(* CODESYS project Syn_Visu_9.4.0.library
   Version: 9.4.0.0
   Title: SynVisu
   Placeholder: SynVisu
   Company: Syntegon Group
   DefaultNamespace: SynVisu

Project tree, tasks and I/O mapping:
  libraries: Tc2_System, * (Beckhoff Automation GmbH)
  DUTs/
    data type E_VisuBodyRole
    data type E_VisuBodyShape
    data type E_VisuCartesianAxes
    data type E_VisuComponentType
    data type E_VisuModuleKind
    data type E_VisuProductShape
    data type E_VisuProductState
    data type ST_VisuBody
    data type ST_VisuBodyState
    data type ST_VisuCartesian
    data type ST_VisuCartesianConfig
    data type ST_VisuCartesianState
    data type ST_VisuConveyor
    data type ST_VisuConveyorConfig
    data type ST_VisuConveyorState
    data type ST_VisuDelta
    data type ST_VisuDeltaConfig
    data type ST_VisuDeltaState
    data type ST_VisuDetector
    data type ST_VisuDetectorConfig
    data type ST_VisuDetectorState
    data type ST_VisuFault
    data type ST_VisuFinger
    data type ST_VisuFingerState
    data type ST_VisuGantryMover
    data type ST_VisuLimitArea
    data type ST_VisuLoopMover
    data type ST_VisuManifest
    data type ST_VisuManifestEntry
    data type ST_VisuPlanarPose
    data type ST_VisuPose
    data type ST_VisuPosition
    data type ST_VisuProduct
    data type ST_VisuProductType
    data type ST_VisuStation
    data type ST_VisuStationConfig
    data type ST_VisuStationState
    data type ST_VisuTrackModule
    data type ST_VisuTrackModuleState
    data type ST_VisuWorkingArea
    data type ST_VisuXtsGantry
    data type ST_VisuXtsGantryConfig
    data type ST_VisuXtsGantryState
    data type ST_VisuXtsLoop
    data type ST_VisuXtsLoopConfig
    data type ST_VisuXtsLoopState
    data type ST_VisuZone
  GVLs/
    global variables VISU_GlobalConst
    global variables VISU_GlobalConst_Param
  POUs/
    function block _FB_VisuBodyComponent [ST]: m_ClearBodies, m_Parts, m_Register, m_SetBody, m_SetBodyActive, m_SetFault, m_SetOriginShift, m_SetPose
    function block _FB_VisuCartesian [ST]: m_ApplyConfig, m_ComponentType, m_Configure, m_Fingers, m_LimitArea, m_SetAxes, m_SetFault, m_SetFingerState, m_SetKinematics, m_SetOriginShift, m_Zones
    function block _FB_VisuComponent [ST]: m_ComponentType, m_DcTime, m_Id, m_NotifyConfigChanged, m_Register, m_SymbolPath
    function block _FB_VisuConveyor [ST]: m_ApplyConfig, m_BeltPosition, m_ComponentType, m_Configure, m_FindProduct, m_GetProduct, m_IndexInsert, m_IndexRebuild, m_IndexSlotOf, m_LatchProduct, m_MoveProduct, m_ProductCount, m_ProductPose, m_RemoveProduct, m_RemoveProductsBeyond, m_SetBeltPosition, m_SetBodyVisible, m_SetFault, m_SetModuloBeltPosition, m_SetOriginShift, m_SetProductState, m_SetProductType, m_StaysInRegister
    function block _FB_VisuDelta [ST]: m_ApplyConfig, m_BasePose, m_ComponentType, m_Configure, m_Fingers, m_LimitArea, m_SetFault, m_SetFingerState, m_SetOriginShift, m_SetTcp, m_SetWorkingArea, m_Zones
    function block _FB_VisuDetector [ST]: m_Parts, m_Zones
    function block _FB_VisuRobot [ST]: m_ClearFingers, m_ClearLimitArea, m_ClearTcpLimitArea, m_Fingers, m_LimitArea, m_SetFinger, m_SetLimitArea, m_SetTcpLimitArea
    function block _FB_VisuSensor [ST]: m_ComponentType, m_Configure, m_SetSignal
    function block _FB_VisuStation [ST]: m_ComponentType, m_Configure, m_Parts, m_Zones
    function block _FB_VisuVision [ST]: m_ComponentType, m_Configure
    function block _FB_VisuXtsGantry [ST]: m_ApplyConfig, m_ComponentType, m_Configure, m_Fingers, m_LimitArea, m_Modules, m_SetFault, m_SetMover, m_SetMoverCount, m_SetOriginShift, m_SetZPosition, m_Zones
    function block _FB_VisuXtsLoop [ST]: m_ApplyConfig, m_ComponentType, m_Configure, m_Fingers, m_LimitArea, m_Modules, m_SetFault, m_SetMover, m_SetMoverCount, m_SetOriginShift, m_Zones
    function block _FB_VisuXtsTrack [ST]: m_ClearModules, m_Modules, m_SetModule, m_SetModuleFault, m_TrackLength
    function block _FB_VisuZoneComponent [ST]: m_ClearZones, m_SetZone, m_Zones
    function _FC_GetVersionSynVisu [ST]
*)

// DUTs/E_VisuBodyRole
{attribute 'qualified_only'}
{attribute 'strict'}
TYPE E_VisuBodyRole :
(
	(* Values are part of the gateway contract: append, never renumber. What a body stands for sets its look. *)
	STRUCTURE := 0,		// machine part: lit, with shadow
	SENSOR := 1,		// sensing part, e.g. a lens or a light barrier head: lit, in its own colour
	BEAM := 2,			// overlay on the zones layer, lights up while active
	FIELD_OF_VIEW := 3	// overlay on the zones layer, lights up while active
) UINT;
END_TYPE

// DUTs/E_VisuBodyShape
{attribute 'qualified_only'}
{attribute 'strict'}
TYPE E_VisuBodyShape :
(
	(* Values are part of the gateway contract: append, never renumber. *)
	BOX := 0,			// box: fLength x fWidth x fHeight
	CYLINDER := 1,		// cylinder: fLength and fWidth are its two diameters
	FRUSTUM := 2		// rectangular pyramid stump: bottom fLength x fWidth, top fTopLength x fTopWidth
) UINT;
END_TYPE

// DUTs/E_VisuCartesianAxes
{attribute 'qualified_only'}
{attribute 'strict'}
TYPE E_VisuCartesianAxes :
(
	(* Values are part of the gateway contract: append, never renumber. Which axes a Cartesian robot has. *)
	XYZ := 0,	// rails along local Y, bridge (Y), carriage (X) and column (Z)
	XZ := 1,	// no Y axis: a fixed beam along local X at fRailHeight, carriage (X) and column (Z); Y is always 0
	XY := 2		// no Z axis: rails, bridge (Y) and carriage (X); the column has a fixed length, the flange stays at fZMin
) UINT;
END_TYPE

// DUTs/E_VisuComponentType
{attribute 'qualified_only'}
{attribute 'strict'}
TYPE E_VisuComponentType :
(
	(* Values are part of the gateway contract: append, never renumber. *)
	NONE := 0,
	CONVEYOR := 1,
	DELTA := 2,
	XTS_GANTRY := 3,
	XTS_LOOP := 4,
	CARTESIAN := 5,
	VISION := 6,
	SENSOR := 7,
	STATION := 8
) UINT;
END_TYPE

// DUTs/E_VisuModuleKind
{attribute 'qualified_only'}
{attribute 'strict'}
TYPE E_VisuModuleKind :
(
	(* Values are part of the gateway contract: append, never renumber. What an XTS track module is. *)
	STRAIGHT := 0,		// straight motor module
	CURVE_LEFT := 1,	// curve module: turns the track by a quarter circle (90 deg) to the left
	CURVE_RIGHT := 2	// curve module: turns the track by a quarter circle (90 deg) to the right
) UINT;
END_TYPE

// DUTs/E_VisuProductShape
{attribute 'qualified_only'}
{attribute 'strict'}
TYPE E_VisuProductShape :
(
	(* Values are part of the gateway contract: append, never renumber. *)
	BOX := 0,			// box: fLength x fWidth x fHeight
	CYLINDER := 1,		// cylinder: fLength and fWidth are its diameters along and across the conveying direction
	ROUNDED_BOX := 2	// box with rounded vertical edges of fCornerRadius (pouches, flow packs)
) UINT;
END_TYPE

// DUTs/E_VisuProductState
{attribute 'qualified_only'}
{attribute 'strict'}
TYPE E_VisuProductState :
(
	(* Values are part of the gateway contract: append, never renumber. *)
	DETECTED := 0,
	ASSIGNED := 1,
	PICKED := 2,
	REJECTED := 3,
	PLACED := 4
) UINT;
END_TYPE

// DUTs/ST_VisuBody
TYPE ST_VisuBody :
STRUCT
	(* One solid a component is drawn from, so the visualisation needs no code of its own for it. It stands on
	   its bottom face and extends along its local +Z. *)
	eShape : E_VisuBodyShape;
	eRole : E_VisuBodyRole;
	stPose : ST_VisuPose; // bottom centre in the component's frame (from its stPose), not MCS
	fLength : LREAL; // mm along the body's local X
	fWidth : LREAL; // mm along the body's local Y
	fHeight : LREAL; // mm along the body's local Z
	fTopLength : LREAL; // mm, top face of a FRUSTUM
	fTopWidth : LREAL; // mm, top face of a FRUSTUM
END_STRUCT
END_TYPE

// DUTs/ST_VisuBodyState
TYPE ST_VisuBodyState :
STRUCT
	bActive : BOOL; // a BEAM or FIELD_OF_VIEW lights up, e.g. an interrupted light barrier
END_STRUCT
END_TYPE

// DUTs/ST_VisuCartesian
TYPE ST_VisuCartesian :
STRUCT
	(* One visualised Cartesian robot. Register the instance's symbol path in the manifest with
	   eType := E_VisuComponentType.CARTESIAN. *)
	stConfig : ST_VisuCartesianConfig; // read at discovery and after nConfigVersion changes
	stState : ST_VisuCartesianState; // read every gateway cycle
END_STRUCT
END_TYPE

// DUTs/ST_VisuCartesianConfig
TYPE ST_VisuCartesianConfig :
STRUCT
	(* Cartesian robot: two fixed rails along local +Y, a bridge travelling in Y, a carriage on it travelling in X
	   and a vertical column (Z) ending at the gripper flange. Local frame: origin at axis X = Y = 0, Z up; the
	   flange is at (X, Y, Z). Without a Y axis (eAxes XZ) a fixed beam along X at fRailHeight replaces rails and
	   bridge and Y is 0; without a Z axis (XY) the column has a fixed length and the flange stays at fZMin. *)
	stPose : ST_VisuPose; // MCS
	eAxes : E_VisuCartesianAxes := E_VisuCartesianAxes.XYZ; // which axes the robot has (set by m_SetKinematics)
	fXMin : LREAL; // mm, X stroke
	fXMax : LREAL; // mm
	fYMin : LREAL; // mm, Y stroke
	fYMax : LREAL; // mm
	fZMin : LREAL; // mm, Z stroke
	fZMax : LREAL; // mm
	fRailHeight : LREAL; // mm, top of the rails above the local origin; the bridge sits on them
	stLimitArea : ST_VisuLimitArea; // optional box in the robot frame that further restricts the working area
	stTcpLimitArea : ST_VisuLimitArea; // optional box around the gripper flange, along the robot frame's axes
	nZoneCount : UINT;
	aZones : ARRAY[0..VISU_GlobalConst_Param.VISU_un_MAX_ZONES - 1] OF ST_VisuZone; // pick and place zones
	nFingerCount : UINT; // 0 = no gripper definition
	aFingers : ARRAY[0..VISU_GlobalConst_Param.VISU_un_MAX_FINGERS - 1] OF ST_VisuFinger;
	(* mm in the local frame from stPose: origin of the robot's coordinate system as shown (origin triad, local
	   measuring coordinates). The geometry and axis values stay relative to stPose. *)
	stOriginShift : ST_VisuPosition;
END_STRUCT
END_TYPE

// DUTs/ST_VisuCartesianState
TYPE ST_VisuCartesianState :
STRUCT
	nTimestamp : ULINT; // DC time of the writing cycle, ns since 2000-01-01 (set by _FB_VisuCartesian)
	fX : LREAL; // mm, actual value: the gripper flange
	fY : LREAL; // mm, actual value
	fZ : LREAL; // mm, actual value
	bGripperActive : BOOL; // used only when no fingers are configured
	aFingerStates : ARRAY[0..VISU_GlobalConst_Param.VISU_un_MAX_FINGERS - 1] OF ST_VisuFingerState; // one per configured finger
	stFault : ST_VisuFault; // fault of the robot (set by _FB_VisuCartesian.m_SetFault)
END_STRUCT
END_TYPE

// DUTs/ST_VisuConveyor
TYPE ST_VisuConveyor :
STRUCT
	(* One visualised conveyor. Register the instance's symbol path in the manifest with
	   eType := E_VisuComponentType.CONVEYOR. *)
	stConfig : ST_VisuConveyorConfig; // read at discovery and after nConfigVersion changes
	stState : ST_VisuConveyorState; // read every gateway cycle
END_STRUCT
END_TYPE

// DUTs/ST_VisuConveyorConfig
TYPE ST_VisuConveyorConfig :
STRUCT
	stPose : ST_VisuPose; // belt start on the belt surface; local +X = conveying direction
	fLength : LREAL; // mm
	fWidth : LREAL; // mm
	nProductTypeCount : UINT;
	aProductTypes : ARRAY[0..VISU_GlobalConst_Param.VISU_un_MAX_PRODUCT_TYPES - 1] OF ST_VisuProductType;
	bBody : BOOL := TRUE; // TRUE = the belt is drawn as a body; FALSE = a conveyor without one (products, zones and axis only)
	(* mm in the local frame from stPose: origin of the conveyor's coordinate system. Belt coordinates (zones'
	   fStart, fEnd, fCcsOffset) count from this origin. 0 = the belt start. *)
	stOriginShift : ST_VisuPosition;
END_STRUCT
END_TYPE

// DUTs/ST_VisuConveyorState
TYPE ST_VisuConveyorState :
STRUCT
	nTimestamp : ULINT; // DC time of the writing cycle, ns since 2000-01-01 (set by _FB_VisuConveyor)
	fBeltPosition : LREAL; // continuous belt surface position, mm, no modulo (see _FB_VisuConveyor.m_SetModuloBeltPosition)
	nProductCount : UINT; // entries [0..nProductCount-1] are evaluated
	aProducts : ARRAY[0..VISU_GlobalConst_Param.VISU_un_MAX_PRODUCTS - 1] OF ST_VisuProduct;
	stFault : ST_VisuFault; // fault of the conveyor (set by _FB_VisuConveyor.m_SetFault)
END_STRUCT
END_TYPE

// DUTs/ST_VisuDelta
TYPE ST_VisuDelta :
STRUCT
	(* One visualised Delta robot. Register the instance's symbol path in the manifest with
	   eType := E_VisuComponentType.DELTA. *)
	stConfig : ST_VisuDeltaConfig; // read at discovery and after nConfigVersion changes
	stState : ST_VisuDeltaState; // read every gateway cycle
END_STRUCT
END_TYPE

// DUTs/ST_VisuDeltaConfig
TYPE ST_VisuDeltaConfig :
STRUCT
	(* Geometry the visualisation uses to derive the arm posture from the TCP.
	   Arm 1 lies along the base's local +X; arms 2 and 3 follow counter-clockwise
	   (seen from above) at 120 deg each. *)
	stPose : ST_VisuPose; // base centre in the MCS
	fBaseRadius : LREAL; // mm, base centre to shoulder joint
	fEffectorRadius : LREAL; // mm, effector centre to lower-arm joint
	fUpperArmLength : LREAL; // mm
	fLowerArmLength : LREAL; // mm
	stWorkingArea : ST_VisuWorkingArea;
	stLimitArea : ST_VisuLimitArea; // optional box that further restricts the working area
	stTcpLimitArea : ST_VisuLimitArea; // optional box around the TCP, relative to it along the robot frame's axes
	nZoneCount : UINT;
	aZones : ARRAY[0..VISU_GlobalConst_Param.VISU_un_MAX_ZONES - 1] OF ST_VisuZone; // pick and place zones
	nFingerCount : UINT; // 0 = no gripper definition
	aFingers : ARRAY[0..VISU_GlobalConst_Param.VISU_un_MAX_FINGERS - 1] OF ST_VisuFinger;
	(* mm in the local frame from stPose: origin of the robot's coordinate system as shown (origin triad, local
	   measuring coordinates). The geometry, working area and limit area stay relative to stPose. *)
	stOriginShift : ST_VisuPosition;
END_STRUCT
END_TYPE

// DUTs/ST_VisuDeltaState
TYPE ST_VisuDeltaState :
STRUCT
	nTimestamp : ULINT; // DC time of the writing cycle, ns since 2000-01-01 (set by _FB_VisuDelta.m_SetTcp)
	stActualTcp : ST_VisuPosition; // MCS, effector centre (the gripper flange); the visualisation derives the arms from it
	stSetpointTcp : ST_VisuPosition; // MCS
	aFingerStates : ARRAY[0..VISU_GlobalConst_Param.VISU_un_MAX_FINGERS - 1] OF ST_VisuFingerState; // one per configured finger
	stFault : ST_VisuFault; // fault of the robot (set by _FB_VisuDelta.m_SetFault)
END_STRUCT
END_TYPE

// DUTs/ST_VisuDetector
TYPE ST_VisuDetector :
STRUCT
	(* One visualised vision system or product sensor. Register the instance's symbol path in the manifest with
	   eType := E_VisuComponentType.VISION or SENSOR; both share this structure. *)
	stConfig : ST_VisuDetectorConfig; // read at discovery and after nConfigVersion changes
	stState : ST_VisuDetectorState; // read every gateway cycle
END_STRUCT
END_TYPE

// DUTs/ST_VisuDetectorConfig
TYPE ST_VisuDetectorConfig :
STRUCT
	(* A detector (vision system, product sensor): its zones on the conveyors and the bodies it is drawn from. *)
	stPose : ST_VisuPose; // MCS; a vision system's lens looking along local -Z, a sensor's head
	nZoneCount : UINT;
	aZones : ARRAY[0..VISU_GlobalConst_Param.VISU_un_MAX_ZONES - 1] OF ST_VisuZone; // where it detects
	nBodyCount : UINT;
	aBodies : ARRAY[0..VISU_GlobalConst_Param.VISU_un_MAX_BODIES - 1] OF ST_VisuBody;
	(* mm in the local frame from stPose: origin of the detector's coordinate system as shown (origin triad, local
	   measuring coordinates). The bodies stay relative to stPose. *)
	stOriginShift : ST_VisuPosition;
END_STRUCT
END_TYPE

// DUTs/ST_VisuDetectorState
TYPE ST_VisuDetectorState :
STRUCT
	nTimestamp : ULINT; // DC time of the writing cycle, ns since 2000-01-01 (set by _FB_VisuDetector)
	aBodyStates : ARRAY[0..VISU_GlobalConst_Param.VISU_un_MAX_BODIES - 1] OF ST_VisuBodyState; // one per configured body
	stFault : ST_VisuFault; // fault of the detector (set by _FB_VisuDetector.m_SetFault)
END_STRUCT
END_TYPE

// DUTs/ST_VisuFault
(* Fault of a component or an XTS mover: drawn red with sMessage while bActive (contract, protocol 8). *)
TYPE ST_VisuFault :
STRUCT
	bActive : BOOL; // TRUE while the fault is active
	sMessage : STRING(80); // shown to the operator; empty shows 'Fault'
END_STRUCT
END_TYPE

// DUTs/ST_VisuFinger
TYPE ST_VisuFinger :
STRUCT
	(* One gripper finger, always drawn as a cylinder. Its frame's origin is the centre of its top face; it extends
	   along its local -Z. The grip point, where a carried product's top touches, is the centre of its bottom face. *)
	fDiameter : LREAL; // mm
	fHeight : LREAL; // mm
END_STRUCT
END_TYPE

// DUTs/ST_VisuFingerState
TYPE ST_VisuFingerState :
STRUCT
	stPose : ST_VisuPose; // MCS, absolute: pose of the finger's frame (centre of its top face)
	bActive : BOOL; // the finger grips
END_STRUCT
END_TYPE

// DUTs/ST_VisuGantryMover
TYPE ST_VisuGantryMover :
STRUCT
	nId : UDINT; // unique within the gantry, > 0; referenced by a carried product's nMoverId
	bValid : BOOL; // invalid entries are not shown
	fPosition : LREAL; // mm along the track (local +Y), actual value
	fX : LREAL; // mm, X axis on the mover, actual value
	bGripperActive : BOOL; // used only when no fingers are configured
	aFingerStates : ARRAY[0..VISU_GlobalConst_Param.VISU_un_MAX_FINGERS - 1] OF ST_VisuFingerState; // one per configured finger
	stFault : ST_VisuFault; // fault of this mover
END_STRUCT
END_TYPE

// DUTs/ST_VisuLimitArea
TYPE ST_VisuLimitArea :
STRUCT
	(* Axis-aligned box along the robot frame's axes (turned with its stPose). As stLimitArea it lies in the robot
	   frame (relative to stPose, the frame its working area is given in) and further restricts the working area, e.g.
	   so that neighbouring robots cannot collide (_FB_VisuRobot.m_SetLimitArea). As stTcpLimitArea it lies around the
	   TCP (XTS gantry: every mover's gripper flange), relative to it, and moves with it without turning
	   (_FB_VisuRobot.m_SetTcpLimitArea): the visualisation flags it when it overlaps another robot's limit area or
	   TCP limit area or leaves its own robot's limit area. Delta, XTS gantry and Cartesian robot; an XTS loop has
	   neither. *)
	fXMin : LREAL; // mm
	fXMax : LREAL; // mm
	fYMin : LREAL; // mm
	fYMax : LREAL; // mm
	fZMin : LREAL; // mm relative to the base or the TCP (below it: negative)
	fZMax : LREAL; // mm relative to the base or the TCP
	bActive : BOOL; // FALSE: no box, nothing is drawn or checked
END_STRUCT
END_TYPE

// DUTs/ST_VisuLoopMover
TYPE ST_VisuLoopMover :
STRUCT
	nId : UDINT; // unique within the loop, > 0; referenced by a carried product's nMoverId
	bValid : BOOL; // invalid entries are not shown
	fPosition : LREAL; // mm along the loop from the start of the lower straight, in the conveying direction
	aFingerStates : ARRAY[0..VISU_GlobalConst_Param.VISU_un_MAX_FINGERS - 1] OF ST_VisuFingerState; // one per configured finger
	stFault : ST_VisuFault; // fault of this mover
END_STRUCT
END_TYPE

// DUTs/ST_VisuManifest
TYPE ST_VisuManifest :
STRUCT
	(* Discovery entry point. The application declares one instance at the fixed symbol
	   GVL_Visu.stManifest; the gateway starts reading there. *)
	nProtocolVersion : UINT := VISU_GlobalConst.VISU_un_PROTOCOL_VERSION;
	(* Increment after any change to the manifest or to a component's stConfig. *)
	nConfigVersion : UDINT := 1;
	nCount : UINT; // entries [0..nCount-1] are evaluated
	aEntries : ARRAY[0..VISU_GlobalConst_Param.VISU_un_MAX_MANIFEST_ENTRIES - 1] OF ST_VisuManifestEntry;
	(* Version of the Syn_Visu library actually running, e.g. '5.1.0', shown by the visualisation. Since 5.1.0;
	   last, so the members before it keep their place. *)
	sLibraryVersion : STRING(15);
END_STRUCT
END_TYPE

// DUTs/ST_VisuManifestEntry
TYPE ST_VisuManifestEntry :
STRUCT
	nId : UDINT; // unique within the manifest, > 0; used for all cross-references
	eType : E_VisuComponentType;
	sName : STRING(80); // display name
	sPath : STRING(255); // symbol path of the ST_VisuConveyor / ST_VisuDelta instance, e.g. 'MAIN.stInfeed'
END_STRUCT
END_TYPE

// DUTs/ST_VisuPlanarPose
TYPE ST_VisuPlanarPose :
STRUCT
	(* Position plus rotation about Z, used for product latch poses (in the conveyor's coordinate system). *)
	fX : LREAL; // mm
	fY : LREAL; // mm
	fZ : LREAL; // mm
	fRz : LREAL; // degrees
END_STRUCT
END_TYPE

// DUTs/ST_VisuPose
TYPE ST_VisuPose :
STRUCT
	(* Pose in the MCS: right-handed, Z up, X in product flow direction.
	   Rotation order R = Rz(fRz) * Ry(fRy) * Rx(fRx). *)
	fX : LREAL; // mm
	fY : LREAL; // mm
	fZ : LREAL; // mm
	fRx : LREAL; // degrees
	fRy : LREAL; // degrees
	fRz : LREAL; // degrees
END_STRUCT
END_TYPE

// DUTs/ST_VisuPosition
TYPE ST_VisuPosition :
STRUCT
	(* A point in the MCS, e.g. a Delta's TCP. *)
	fX : LREAL; // mm
	fY : LREAL; // mm
	fZ : LREAL; // mm
END_STRUCT
END_TYPE

// DUTs/ST_VisuProduct
TYPE ST_VisuProduct :
STRUCT
	nId : UDINT;
	bValid : BOOL; // invalid entries are not shown
	stLatchPose : ST_VisuPlanarPose; // conveyor coordinate system (stPose + stOriginShift), bottom centre at latch time
	fLatchBeltPosition : LREAL; // conveyor fBeltPosition at latch time, mm
	eState : E_VisuProductState;
	ePreviousState : E_VisuProductState; // state before the last change; equals eState until the first change
	(* Manifest id of the client that made the last change: the detector or station that latched it, the robot it
	   is assigned to, picked by or placed by, the station that rejected it; 0 = none given. *)
	nLastClientId : UDINT;
	nMoverId : UDINT; // mover of an XTS gantry or loop carrying the product, 0 = none
	nFingerId : UDINT; // gripper finger (1-based) the product hangs from while picked, 0 = the gripper flange
	nProductType : UDINT; // id in the conveyor's aProductTypes
END_STRUCT
END_TYPE

// DUTs/ST_VisuProductType
TYPE ST_VisuProductType :
STRUCT
	nId : UDINT;
	fLength : LREAL; // mm, along the conveying direction
	fWidth : LREAL; // mm
	fHeight : LREAL; // mm
	eShape : E_VisuProductShape; // solid of the product
	fCornerRadius : LREAL; // mm, rounded vertical edges of a ROUNDED_BOX
END_STRUCT
END_TYPE

// DUTs/ST_VisuStation
TYPE ST_VisuStation :
STRUCT
	(* One visualised station. Register the instance's symbol path in the manifest with
	   eType := E_VisuComponentType.STATION. *)
	stConfig : ST_VisuStationConfig; // read at discovery and after nConfigVersion changes
	stState : ST_VisuStationState; // read every gateway cycle
END_STRUCT
END_TYPE

// DUTs/ST_VisuStationConfig
TYPE ST_VisuStationConfig :
STRUCT
	(* A station (reject unit, labeller, printer, check weigher): its zones on the conveyors and the bodies it is
	   drawn from. *)
	stPose : ST_VisuPose; // MCS, the station's origin; its bodies are placed relative to it
	nZoneCount : UINT;
	aZones : ARRAY[0..VISU_GlobalConst_Param.VISU_un_MAX_ZONES - 1] OF ST_VisuZone; // where it works on products
	nBodyCount : UINT;
	aBodies : ARRAY[0..VISU_GlobalConst_Param.VISU_un_MAX_BODIES - 1] OF ST_VisuBody;
	(* mm in the local frame from stPose: origin of the station's coordinate system as shown (origin triad, local
	   measuring coordinates). The bodies stay relative to stPose. *)
	stOriginShift : ST_VisuPosition;
END_STRUCT
END_TYPE

// DUTs/ST_VisuStationState
TYPE ST_VisuStationState :
STRUCT
	nTimestamp : ULINT; // DC time of the writing cycle, ns since 2000-01-01 (set by _FB_VisuStation)
	aBodyStates : ARRAY[0..VISU_GlobalConst_Param.VISU_un_MAX_BODIES - 1] OF ST_VisuBodyState; // one per configured body; an active body lights up
	stFault : ST_VisuFault; // fault of the station (set by _FB_VisuStation.m_SetFault)
END_STRUCT
END_TYPE

// DUTs/ST_VisuTrackModule
TYPE ST_VisuTrackModule :
STRUCT
	(* One XTS motor module of a track, in the order the movers run along it. Each module starts where the one
	   before it ends; a curve module is drawn as a quarter circle as long as fLength. *)
	eKind : E_VisuModuleKind;
	fLength : LREAL; // mm along the track (track positions), VISU_GlobalConst.VISU_lr_XTS_MODULE_LENGTH for an XTS module
END_STRUCT
END_TYPE

// DUTs/ST_VisuTrackModuleState
TYPE ST_VisuTrackModuleState :
STRUCT
	stFault : ST_VisuFault; // fault of this track module (set by _FB_VisuXtsTrack.m_SetModuleFault)
END_STRUCT
END_TYPE

// DUTs/ST_VisuWorkingArea
TYPE ST_VisuWorkingArea :
STRUCT
	(* Limit shape the PLC enforces: vertical cylinder in the robot frame, optional cone below. *)
	fRadius : LREAL; // mm
	fZMin : LREAL; // mm relative to the base (below the base: negative)
	fZMax : LREAL; // mm relative to the base
	fConeHeight : LREAL; // mm below fZMin; 0 = no cone
	fConeBottomRadius : LREAL; // mm
END_STRUCT
END_TYPE

// DUTs/ST_VisuXtsGantry
TYPE ST_VisuXtsGantry :
STRUCT
	(* One visualised XTS gantry (e.g. IDH). Register the instance's symbol path in the manifest with
	   eType := E_VisuComponentType.XTS_GANTRY. *)
	stConfig : ST_VisuXtsGantryConfig; // read at discovery and after nConfigVersion changes
	stState : ST_VisuXtsGantryState; // read every gateway cycle
END_STRUCT
END_TYPE

// DUTs/ST_VisuXtsGantryConfig
TYPE ST_VisuXtsGantryConfig :
STRUCT
	(* Straight XTS track of track modules, carried by a common Z axis; every mover carries an X axis with a
	   gripper flange at its end. Local frame: origin at the track start on top of the movers with Z = 0; the track runs
	   along local +Y, the X axes along local +X, the Z axis along local +Z (up). *)
	stPose : ST_VisuPose; // MCS
	nModuleCount : UINT; // entries [0..nModuleCount-1] are evaluated
	aModules : ARRAY[0..VISU_GlobalConst_Param.VISU_un_MAX_MODULES - 1] OF ST_VisuTrackModule; // from the track start along local +Y
	fXMin : LREAL; // mm, X stroke
	fXMax : LREAL; // mm
	fZMin : LREAL; // mm, Z stroke
	fZMax : LREAL; // mm
	fToolOffsetX : LREAL; // mm, gripper flange ahead of the X axis zero along local +X
	fToolOffsetZ : LREAL; // mm, gripper flange relative to the mover top (below: negative)
	fMoverLength : LREAL; // mm, along the track
	fMoverWidth : LREAL; // mm
	stLimitArea : ST_VisuLimitArea; // optional box in the gantry frame that further restricts the working area
	stTcpLimitArea : ST_VisuLimitArea; // optional box around every mover's gripper flange, along the gantry frame's axes
	nZoneCount : UINT;
	aZones : ARRAY[0..VISU_GlobalConst_Param.VISU_un_MAX_ZONES - 1] OF ST_VisuZone; // pick and place zones
	nFingerCount : UINT; // fingers of every mover's gripper, 0 = no gripper definition
	aFingers : ARRAY[0..VISU_GlobalConst_Param.VISU_un_MAX_FINGERS - 1] OF ST_VisuFinger;
	(* mm in the local frame from stPose: origin of the gantry's coordinate system as shown (origin triad, local
	   measuring coordinates). The geometry and mover positions stay relative to stPose. *)
	stOriginShift : ST_VisuPosition;
END_STRUCT
END_TYPE

// DUTs/ST_VisuXtsGantryState
TYPE ST_VisuXtsGantryState :
STRUCT
	nTimestamp : ULINT; // DC time of the writing cycle, ns since 2000-01-01 (set by _FB_VisuXtsGantry)
	fZ : LREAL; // mm, common Z axis, actual value
	nMoverCount : UINT; // entries [0..nMoverCount-1] are evaluated
	aMovers : ARRAY[0..VISU_GlobalConst_Param.VISU_un_MAX_MOVERS - 1] OF ST_VisuGantryMover;
	aModuleStates : ARRAY[0..VISU_GlobalConst_Param.VISU_un_MAX_MODULES - 1] OF ST_VisuTrackModuleState; // index as in stConfig.aModules
	stFault : ST_VisuFault; // fault of the whole gantry (set by _FB_VisuXtsGantry.m_SetFault)
END_STRUCT
END_TYPE

// DUTs/ST_VisuXtsLoop
TYPE ST_VisuXtsLoop :
STRUCT
	(* One visualised XTS loop (e.g. Fxx). Register the instance's symbol path in the manifest with
	   eType := E_VisuComponentType.XTS_LOOP. *)
	stConfig : ST_VisuXtsLoopConfig; // read at discovery and after nConfigVersion changes
	stState : ST_VisuXtsLoopState; // read every gateway cycle
END_STRUCT
END_TYPE

// DUTs/ST_VisuXtsLoopConfig
TYPE ST_VisuXtsLoopConfig :
STRUCT
	(* Closed XTS loop of track modules standing in the local X-Z plane, e.g. two straights joined at each end by two
	   CURVE_LEFT modules. Local frame: origin at the start of the first module, which runs along local +X in the
	   conveying direction; a left curve turns up towards +Z. *)
	stPose : ST_VisuPose; // MCS
	nModuleCount : UINT; // entries [0..nModuleCount-1] are evaluated
	aModules : ARRAY[0..VISU_GlobalConst_Param.VISU_un_MAX_MODULES - 1] OF ST_VisuTrackModule; // the chain should end where it starts
	fToolOffset : LREAL; // mm, gripper flange (tool point) of a mover outwards from the track
	fMoverLength : LREAL; // mm, along the track
	fMoverWidth : LREAL; // mm
	nZoneCount : UINT;
	aZones : ARRAY[0..VISU_GlobalConst_Param.VISU_un_MAX_ZONES - 1] OF ST_VisuZone; // pick and place zones
	nFingerCount : UINT; // fingers of every mover's gripper, 0 = no gripper definition
	aFingers : ARRAY[0..VISU_GlobalConst_Param.VISU_un_MAX_FINGERS - 1] OF ST_VisuFinger;
	(* mm in the local frame from stPose: origin of the loop's coordinate system as shown (origin triad, local
	   measuring coordinates). The geometry and mover positions stay relative to stPose. *)
	stOriginShift : ST_VisuPosition;
END_STRUCT
END_TYPE

// DUTs/ST_VisuXtsLoopState
TYPE ST_VisuXtsLoopState :
STRUCT
	nTimestamp : ULINT; // DC time of the writing cycle, ns since 2000-01-01 (set by _FB_VisuXtsLoop)
	nMoverCount : UINT; // entries [0..nMoverCount-1] are evaluated
	aMovers : ARRAY[0..VISU_GlobalConst_Param.VISU_un_MAX_MOVERS - 1] OF ST_VisuLoopMover;
	aModuleStates : ARRAY[0..VISU_GlobalConst_Param.VISU_un_MAX_MODULES - 1] OF ST_VisuTrackModuleState; // index as in stConfig.aModules
	stFault : ST_VisuFault; // fault of the whole loop (set by _FB_VisuXtsLoop.m_SetFault)
END_STRUCT
END_TYPE

// DUTs/ST_VisuZone
TYPE ST_VisuZone :
STRUCT
	(* A stretch of a conveyor that belongs to a component: where a robot picks or places, where a detector
	   detects. The visualisation draws every zone alike; fStart = fEnd is a line across the belt. *)
	nConveyorId : UDINT; // manifest id of the conveyor
	fStart : LREAL; // mm along the conveyor's local X (belt coordinates, not MCS)
	fEnd : LREAL; // mm along the conveyor's local X
	(* mm before fEnd, against the conveying direction: the robot may allocate products in the zone only up to
	   fEnd - fAllocationOffset, so it does not move out of the zone while approaching. 0 = no allocation limit. *)
	fAllocationOffset : LREAL;
	(* mm along the conveyor's local X, like fStart / fEnd: position of the robot's conveyor coordinate system (CCS)
	   on this conveyor. Drawn as a solid line across the zone; may lie outside the zone, but on the belt. *)
	fCcsOffset : LREAL;
	(* mm along the conveyor's local Y (from its origin, like the products' latch pose): the zone's sides across
	   the belt, in any order. fStartY = fEndY = the whole belt width. Clipped to the belt when drawn. *)
	fStartY : LREAL;
	fEndY : LREAL;
END_STRUCT
END_TYPE

// GVLs/VISU_GlobalConst
(****************************************************************************************************<br>
© Syntegon Group.<br>
All rights reserved, also regarding any disposal, exploitation, reproduction, editing, distribution,<br>
as well as in the event of applications for industrial property rights.<br>
*****************************************************************************************************<br>
DESCRIPTION:<br>
Global constants of the Syn_Visu library.<br>
****************************************************************************************************)
{attribute 'qualified_only'}
VAR_GLOBAL CONSTANT
	(* Version of the PLC <-> gateway contract. The gateway refuses to read a PLC whose manifest
	   reports a different value. Bump together with PROTOCOL_VERSION in the gateway.
	   2: the Delta reports only its TCP; the visualisation derives the arm posture.
	   3: work area renamed to working area, windows to zones.
	   4: XTS gantry and XTS loop, product nMoverId, fEncoder renamed to fBeltPosition.
	   5: Cartesian robot.
	   6: Delta limit area, zone allocation offset.
	   7: gripper fingers; tool rotations (Delta rz, IDH C, Cartesian C/A and tool length) removed.
	   8: faults of components and XTS movers (stFault).
	   9: zone fCcsOffset, stOriginShift in every config.
	   10: product type eShape and fCornerRadius.
	   11: zones without kind, product nDetectorId, vision system and product sensor (ST_VisuDetector).
	   12: XTS tracks as chains of track modules (straight, quarter curves) with a fault per module.
	   13: product nLastClientId and ePreviousState instead of nRobotId and nDetectorId; station (ST_VisuStation).
	   14: product stLatchPose in the conveyor's coordinate system instead of the MCS.
	   15: zone fStartY and fEndY, the zone's sides across the belt.
	   16: conveyor bBody, a conveyor may have no body.
	   17: Cartesian robot eAxes (E_VisuCartesianAxes): X, Y, Z or without the Y or the Z axis.
	   18: stLimitArea for the XTS gantry and the Cartesian robot too, not only the Delta.
	   19: stTcpLimitArea, a box around the TCP, for the Delta, the XTS gantry and the Cartesian robot. *)
	VISU_un_PROTOCOL_VERSION			: UINT := 19;
	(* Version of this library as the visualisation shows it (manifest sLibraryVersion). Bump together with
	   _FC_GetVersionSynVisu and the project version. *)
	VISU_str_LIBRARY_VERSION			: STRING(15) := '9.4.0';
	VISU_lr_DEG_TO_RAD					: LREAL := 0.017453292519943295;	// [rad/deg] pi / 180
	VISU_lr_XTS_MODULE_LENGTH			: LREAL := 250;	// [mm] length of an XTS motor module along the track, straight or curve
END_VAR

// GVLs/VISU_GlobalConst_Param
(****************************************************************************************************<br>
© Syntegon Group.<br>
All rights reserved, also regarding any disposal, exploitation, reproduction, editing, distribution,<br>
as well as in the event of applications for industrial property rights.<br>
*****************************************************************************************************<br>
DESCRIPTION:<br>
Library parameters of Syn_Visu: array sizes of the interface structures.<br>
****************************************************************************************************)
{attribute 'qualified_only'}
VAR_GLOBAL CONSTANT
	VISU_un_MAX_MANIFEST_ENTRIES		: UINT := 32;	// [-] components in the manifest
	VISU_un_MAX_PRODUCTS				: UINT := 4800;	// [-] products per conveyor
	VISU_un_PRODUCT_INDEX_SIZE			: UINT := 16384;	// [-] slots of a conveyor's product index by id: a power of two, at least twice VISU_un_MAX_PRODUCTS
	VISU_un_MAX_PRODUCT_TYPES			: UINT := 8;	// [-] product types per conveyor
	VISU_un_MAX_ZONES					: UINT := 8;	// [-] zones per robot or detector
	VISU_un_MAX_MOVERS					: UINT := 40;	// [-] movers per XTS gantry or loop
	VISU_un_MAX_FINGERS					: UINT := 8;	// [-] fingers per gripper
	VISU_un_MAX_BODIES					: UINT := 16;	// [-] bodies per detector
	VISU_un_MAX_MODULES					: UINT := 64;	// [-] track modules per XTS gantry or loop
	VISU_un_INSTANCE_PATH_SKIP			: UINT := 2;	// [-] leading segments of an instance path that are not part of its symbol path: TwinCAT project and PLC project
END_VAR

// POUs/_FB_VisuBodyComponent
(****************************************************************************************************<br>
© Syntegon Group.<br>
All rights reserved, also regarding any disposal, exploitation, reproduction, editing, distribution,<br>
as well as in the event of applications for industrial property rights.<br>
*****************************************************************************************************<br>
DESCRIPTION:<br>
Base of every component drawn from the bodies it describes, with zones on conveyors: detectors<br>
(_FB_VisuVision, _FB_VisuSensor) and stations (_FB_VisuStation). The visualisation needs no code of its<br>
own for them. Bodies: m_SetBody, m_SetBodyActive, m_ClearBodies; also the fault (m_SetFault) and the<br>
origin shift (m_SetOriginShift). m_Register, called every cycle, also stamps the state. A derived FB<br>
tells where these lie in its contract structure through m_Parts. Not used directly.<br>
*****************************************************************************************************<br>
VERSION         ¦ DATE       ¦ NAME      ¦ CHANGE<br>
Syn_Visu 6.0.0  ¦ 2026-11-01 ¦ J.Willner ¦ New: body handling of _FB_VisuDetector, shared with stations<br>
****************************************************************************************************)
FUNCTION_BLOCK ABSTRACT _FB_VisuBodyComponent EXTENDS _FB_VisuZoneComponent

(****************************************************************************************************<br>
© Syntegon Group.<br>
All rights reserved, also regarding any disposal, exploitation, reproduction, editing, distribution,<br>
as well as in the event of applications for industrial property rights.<br>
*****************************************************************************************************<br>
DESCRIPTION:<br>
Removes all bodies, also those m_Configure described. TRUE if there were any.<br>
****************************************************************************************************)
METHOD m_ClearBodies : BOOL
VAR
	p_TempPose							: POINTER TO ST_VisuPose;
	p_TempShift							: POINTER TO ST_VisuPosition;
	p_TempCount							: POINTER TO UINT;
	p_TempBodies						: POINTER TO ARRAY[0..VISU_GlobalConst_Param.VISU_un_MAX_BODIES - 1] OF ST_VisuBody;
	p_TempStates						: POINTER TO ARRAY[0..VISU_GlobalConst_Param.VISU_un_MAX_BODIES - 1] OF ST_VisuBodyState;
	p_TempTimestamp						: POINTER TO ULINT;
	p_TempFault							: POINTER TO ST_VisuFault;
	TempEmpty							: ST_VisuBody;
	un_TempIndex						: UINT;
END_VAR
m_ClearBodies := FALSE;
m_Parts(vo_p_Pose => p_TempPose, vo_p_OriginShift => p_TempShift, vo_p_BodyCount => p_TempCount,
	vo_p_Bodies => p_TempBodies, vo_p_BodyStates => p_TempStates, vo_p_Timestamp => p_TempTimestamp,
	vo_p_Fault => p_TempFault);
IF p_TempCount = 0 OR p_TempBodies = 0 OR p_TempStates = 0 THEN
	RETURN;
END_IF
m_ClearBodies := p_TempCount^ > 0;
FOR un_TempIndex := 0 TO VISU_GlobalConst_Param.VISU_un_MAX_BODIES - 1 DO
	p_TempBodies^[un_TempIndex] := TempEmpty;
	p_TempStates^[un_TempIndex].bActive := FALSE;
END_FOR
p_TempCount^ := 0;
IF m_ClearBodies THEN
	m_NotifyConfigChanged();
END_IF
END_METHOD

(****************************************************************************************************<br>
© Syntegon Group.<br>
All rights reserved, also regarding any disposal, exploitation, reproduction, editing, distribution,<br>
as well as in the event of applications for industrial property rights.<br>
*****************************************************************************************************<br>
DESCRIPTION:<br>
Where the pose, origin shift, bodies, body states, timestamp and fault lie in the derived FB's contract<br>
structure (stConfig.stPose, stConfig.stOriginShift, stConfig.nBodyCount, stConfig.aBodies,<br>
stState.aBodyStates, stState.nTimestamp, stState.stFault).<br>
****************************************************************************************************)
METHOD PROTECTED ABSTRACT m_Parts : BOOL
VAR_OUTPUT
	vo_p_Pose							: POINTER TO ST_VisuPose;
	vo_p_OriginShift					: POINTER TO ST_VisuPosition;
	vo_p_BodyCount						: POINTER TO UINT;
	vo_p_Bodies							: POINTER TO ARRAY[0..VISU_GlobalConst_Param.VISU_un_MAX_BODIES - 1] OF ST_VisuBody;
	vo_p_BodyStates						: POINTER TO ARRAY[0..VISU_GlobalConst_Param.VISU_un_MAX_BODIES - 1] OF ST_VisuBodyState;
	vo_p_Timestamp						: POINTER TO ULINT;
	vo_p_Fault							: POINTER TO ST_VisuFault;
END_VAR
END_METHOD

(****************************************************************************************************<br>
© Syntegon Group.<br>
All rights reserved, also regarding any disposal, exploitation, reproduction, editing, distribution,<br>
as well as in the event of applications for industrial property rights.<br>
*****************************************************************************************************<br>
DESCRIPTION:<br>
As _FB_VisuComponent.m_Register; since such a component may have no cyclic value of its own to report,<br>
this call, made every cycle, also stamps its state with the cycle's DC time.<br>
*****************************************************************************************************<br>
OUTPUT VALUES:<br>
FALSE for vi_udn_Id = 0, an id already used by a different entry, or a full manifest.<br>
****************************************************************************************************)
METHOD m_Register : BOOL
VAR_IN_OUT
	vio_Manifest						: ST_VisuManifest;	// GVL_Visu.stManifest of the application
END_VAR
VAR_INPUT
	vi_udn_Id							: UDINT;	// [-] unique, > 0
	vi_str_Name							: STRING(80);	// display name
END_VAR
VAR
	p_TempPose							: POINTER TO ST_VisuPose;
	p_TempShift							: POINTER TO ST_VisuPosition;
	p_TempCount							: POINTER TO UINT;
	p_TempBodies						: POINTER TO ARRAY[0..VISU_GlobalConst_Param.VISU_un_MAX_BODIES - 1] OF ST_VisuBody;
	p_TempStates						: POINTER TO ARRAY[0..VISU_GlobalConst_Param.VISU_un_MAX_BODIES - 1] OF ST_VisuBodyState;
	p_TempTimestamp						: POINTER TO ULINT;
	p_TempFault							: POINTER TO ST_VisuFault;
END_VAR
m_Register := SUPER^.m_Register(vio_Manifest := vio_Manifest, vi_udn_Id := vi_udn_Id, vi_str_Name := vi_str_Name);
m_Parts(vo_p_Pose => p_TempPose, vo_p_OriginShift => p_TempShift, vo_p_BodyCount => p_TempCount,
	vo_p_Bodies => p_TempBodies, vo_p_BodyStates => p_TempStates, vo_p_Timestamp => p_TempTimestamp,
	vo_p_Fault => p_TempFault);
IF p_TempTimestamp <> 0 THEN
	p_TempTimestamp^ := m_DcTime();
END_IF
END_METHOD

(****************************************************************************************************<br>
© Syntegon Group.<br>
All rights reserved, also regarding any disposal, exploitation, reproduction, editing, distribution,<br>
as well as in the event of applications for industrial property rights.<br>
*****************************************************************************************************<br>
DESCRIPTION:<br>
Describes body vi_un_Body (1-based), a solid the component is drawn from: standing on its bottom centre<br>
vi_Pose in the component's frame and extending along its local +Z. The body count grows to vi_un_Body.<br>
m_Configure of _FB_VisuVision and _FB_VisuSensor sets the first bodies; further ones may be added,<br>
e.g. a bracket. A station describes all of its bodies with this. TRUE if set; the config version only<br>
changes when a value does.<br>
*****************************************************************************************************<br>
OUTPUT VALUES:<br>
FALSE outside 1..VISU_GlobalConst_Param.VISU_un_MAX_BODIES.<br>
****************************************************************************************************)
METHOD m_SetBody : BOOL
VAR_INPUT
	vi_un_Body							: UINT;	// [-] 1-based
	vi_e_Shape							: E_VisuBodyShape;
	vi_e_Role							: E_VisuBodyRole;	// sets its look
	vi_Pose								: ST_VisuPose;	// bottom centre in the component's frame, not MCS
	vi_lr_Length						: LREAL;	// [mm] along the body's local X; a cylinder's diameter
	vi_lr_Width							: LREAL;	// [mm] along the body's local Y; a cylinder's diameter
	vi_lr_Height						: LREAL;	// [mm] along the body's local Z
	vi_lr_TopLength						: LREAL;	// [mm] top face of a FRUSTUM, 0 for other shapes
	vi_lr_TopWidth						: LREAL;	// [mm] top face of a FRUSTUM, 0 for other shapes
END_VAR
VAR
	p_TempPose							: POINTER TO ST_VisuPose;
	p_TempShift							: POINTER TO ST_VisuPosition;
	p_TempCount							: POINTER TO UINT;
	p_TempBodies						: POINTER TO ARRAY[0..VISU_GlobalConst_Param.VISU_un_MAX_BODIES - 1] OF ST_VisuBody;
	p_TempStates						: POINTER TO ARRAY[0..VISU_GlobalConst_Param.VISU_un_MAX_BODIES - 1] OF ST_VisuBodyState;
	p_TempTimestamp						: POINTER TO ULINT;
	p_TempFault							: POINTER TO ST_VisuFault;
	b_TempChanged						: BOOL;
END_VAR
m_SetBody := FALSE;
IF vi_un_Body = 0 OR vi_un_Body > VISU_GlobalConst_Param.VISU_un_MAX_BODIES THEN
	RETURN;
END_IF
m_Parts(vo_p_Pose => p_TempPose, vo_p_OriginShift => p_TempShift, vo_p_BodyCount => p_TempCount,
	vo_p_Bodies => p_TempBodies, vo_p_BodyStates => p_TempStates, vo_p_Timestamp => p_TempTimestamp,
	vo_p_Fault => p_TempFault);
IF p_TempCount = 0 OR p_TempBodies = 0 THEN
	RETURN;
END_IF

(* Member by member: a memory compare would also see the padding of the structure. *)
b_TempChanged := vi_un_Body > p_TempCount^
	OR p_TempBodies^[vi_un_Body - 1].eShape <> vi_e_Shape
	OR p_TempBodies^[vi_un_Body - 1].eRole <> vi_e_Role
	OR Tc2_System.MEMCMP(ADR(p_TempBodies^[vi_un_Body - 1].stPose), ADR(vi_Pose), SIZEOF(vi_Pose)) <> 0
	OR p_TempBodies^[vi_un_Body - 1].fLength <> vi_lr_Length
	OR p_TempBodies^[vi_un_Body - 1].fWidth <> vi_lr_Width
	OR p_TempBodies^[vi_un_Body - 1].fHeight <> vi_lr_Height
	OR p_TempBodies^[vi_un_Body - 1].fTopLength <> vi_lr_TopLength
	OR p_TempBodies^[vi_un_Body - 1].fTopWidth <> vi_lr_TopWidth;
IF b_TempChanged THEN
	p_TempBodies^[vi_un_Body - 1].eShape := vi_e_Shape;
	p_TempBodies^[vi_un_Body - 1].eRole := vi_e_Role;
	p_TempBodies^[vi_un_Body - 1].stPose := vi_Pose;
	p_TempBodies^[vi_un_Body - 1].fLength := vi_lr_Length;
	p_TempBodies^[vi_un_Body - 1].fWidth := vi_lr_Width;
	p_TempBodies^[vi_un_Body - 1].fHeight := vi_lr_Height;
	p_TempBodies^[vi_un_Body - 1].fTopLength := vi_lr_TopLength;
	p_TempBodies^[vi_un_Body - 1].fTopWidth := vi_lr_TopWidth;
	p_TempCount^ := MAX(p_TempCount^, vi_un_Body);
	m_NotifyConfigChanged();
END_IF
m_SetBody := TRUE;
END_METHOD

(****************************************************************************************************<br>
© Syntegon Group.<br>
All rights reserved, also regarding any disposal, exploitation, reproduction, editing, distribution,<br>
as well as in the event of applications for industrial property rights.<br>
*****************************************************************************************************<br>
DESCRIPTION:<br>
Reports whether body vi_un_Body (1-based) is active: it then lights up, e.g. an interrupted beam, a field<br>
of view while the camera triggers, a reject unit's pusher while it rejects. Also stamps the state with the<br>
cycle's DC time.<br>
*****************************************************************************************************<br>
OUTPUT VALUES:<br>
FALSE outside 1..VISU_GlobalConst_Param.VISU_un_MAX_BODIES.<br>
****************************************************************************************************)
METHOD m_SetBodyActive : BOOL
VAR_INPUT
	vi_un_Body							: UINT;	// [-] 1-based
	vi_b_Active							: BOOL;
END_VAR
VAR
	p_TempPose							: POINTER TO ST_VisuPose;
	p_TempShift							: POINTER TO ST_VisuPosition;
	p_TempCount							: POINTER TO UINT;
	p_TempBodies						: POINTER TO ARRAY[0..VISU_GlobalConst_Param.VISU_un_MAX_BODIES - 1] OF ST_VisuBody;
	p_TempStates						: POINTER TO ARRAY[0..VISU_GlobalConst_Param.VISU_un_MAX_BODIES - 1] OF ST_VisuBodyState;
	p_TempTimestamp						: POINTER TO ULINT;
	p_TempFault							: POINTER TO ST_VisuFault;
END_VAR
m_SetBodyActive := FALSE;
IF vi_un_Body = 0 OR vi_un_Body > VISU_GlobalConst_Param.VISU_un_MAX_BODIES THEN
	RETURN;
END_IF
m_Parts(vo_p_Pose => p_TempPose, vo_p_OriginShift => p_TempShift, vo_p_BodyCount => p_TempCount,
	vo_p_Bodies => p_TempBodies, vo_p_BodyStates => p_TempStates, vo_p_Timestamp => p_TempTimestamp,
	vo_p_Fault => p_TempFault);
IF p_TempStates = 0 OR p_TempTimestamp = 0 THEN
	RETURN;
END_IF
p_TempStates^[vi_un_Body - 1].bActive := vi_b_Active;
p_TempTimestamp^ := m_DcTime();
m_SetBodyActive := TRUE;
END_METHOD

(****************************************************************************************************<br>
© Syntegon Group.<br>
All rights reserved, also regarding any disposal, exploitation, reproduction, editing, distribution,<br>
as well as in the event of applications for industrial property rights.<br>
*****************************************************************************************************<br>
DESCRIPTION:<br>
Sets or clears the fault of the component: drawn red with the message while active. The fault stays until<br>
it is cleared with m_SetFault(vi_b_Active := FALSE, vi_str_Message := ''). TRUE if set.<br>
****************************************************************************************************)
METHOD m_SetFault : BOOL
VAR_INPUT
	vi_b_Active							: BOOL;	// TRUE: fault active
	vi_str_Message						: STRING(80);	// shown to the operator; empty shows 'Fault'
END_VAR
VAR
	p_TempPose							: POINTER TO ST_VisuPose;
	p_TempShift							: POINTER TO ST_VisuPosition;
	p_TempCount							: POINTER TO UINT;
	p_TempBodies						: POINTER TO ARRAY[0..VISU_GlobalConst_Param.VISU_un_MAX_BODIES - 1] OF ST_VisuBody;
	p_TempStates						: POINTER TO ARRAY[0..VISU_GlobalConst_Param.VISU_un_MAX_BODIES - 1] OF ST_VisuBodyState;
	p_TempTimestamp						: POINTER TO ULINT;
	p_TempFault							: POINTER TO ST_VisuFault;
END_VAR
m_SetFault := FALSE;
m_Parts(vo_p_Pose => p_TempPose, vo_p_OriginShift => p_TempShift, vo_p_BodyCount => p_TempCount,
	vo_p_Bodies => p_TempBodies, vo_p_BodyStates => p_TempStates, vo_p_Timestamp => p_TempTimestamp,
	vo_p_Fault => p_TempFault);
IF p_TempFault = 0 THEN
	RETURN;
END_IF
p_TempFault^.bActive := vi_b_Active;
p_TempFault^.sMessage := vi_str_Message;
m_SetFault := TRUE;
END_METHOD

(****************************************************************************************************<br>
© Syntegon Group.<br>
All rights reserved, also regarding any disposal, exploitation, reproduction, editing, distribution,<br>
as well as in the event of applications for industrial property rights.<br>
*****************************************************************************************************<br>
DESCRIPTION:<br>
Moves the component's shown coordinate system (origin triad, local measuring coordinates) away from its<br>
pose, in its local frame. The bodies stay relative to the pose. TRUE if anything changed.<br>
****************************************************************************************************)
METHOD m_SetOriginShift : BOOL
VAR_INPUT
	vi_lr_X								: LREAL;	// [mm] along the component's local X
	vi_lr_Y								: LREAL;	// [mm] along the component's local Y, 0 = none
	vi_lr_Z								: LREAL;	// [mm] along the component's local Z, 0 = none
END_VAR
VAR
	p_TempPose							: POINTER TO ST_VisuPose;
	p_TempShift							: POINTER TO ST_VisuPosition;
	p_TempCount							: POINTER TO UINT;
	p_TempBodies						: POINTER TO ARRAY[0..VISU_GlobalConst_Param.VISU_un_MAX_BODIES - 1] OF ST_VisuBody;
	p_TempStates						: POINTER TO ARRAY[0..VISU_GlobalConst_Param.VISU_un_MAX_BODIES - 1] OF ST_VisuBodyState;
	p_TempTimestamp						: POINTER TO ULINT;
	p_TempFault							: POINTER TO ST_VisuFault;
END_VAR
m_SetOriginShift := FALSE;
m_Parts(vo_p_Pose => p_TempPose, vo_p_OriginShift => p_TempShift, vo_p_BodyCount => p_TempCount,
	vo_p_Bodies => p_TempBodies, vo_p_BodyStates => p_TempStates, vo_p_Timestamp => p_TempTimestamp,
	vo_p_Fault => p_TempFault);
IF p_TempShift = 0 THEN
	RETURN;
END_IF
m_SetOriginShift := p_TempShift^.fX <> vi_lr_X OR p_TempShift^.fY <> vi_lr_Y OR p_TempShift^.fZ <> vi_lr_Z;
IF m_SetOriginShift THEN
	p_TempShift^.fX := vi_lr_X;
	p_TempShift^.fY := vi_lr_Y;
	p_TempShift^.fZ := vi_lr_Z;
	m_NotifyConfigChanged();
END_IF
END_METHOD

(****************************************************************************************************<br>
© Syntegon Group.<br>
All rights reserved, also regarding any disposal, exploitation, reproduction, editing, distribution,<br>
as well as in the event of applications for industrial property rights.<br>
*****************************************************************************************************<br>
DESCRIPTION:<br>
Sets the component's pose, for m_Configure of the derived FB. TRUE if it changed.<br>
****************************************************************************************************)
METHOD PROTECTED m_SetPose : BOOL
VAR_INPUT
	vi_Pose								: ST_VisuPose;	// MCS
END_VAR
VAR
	p_TempPose							: POINTER TO ST_VisuPose;
	p_TempShift							: POINTER TO ST_VisuPosition;
	p_TempCount							: POINTER TO UINT;
	p_TempBodies						: POINTER TO ARRAY[0..VISU_GlobalConst_Param.VISU_un_MAX_BODIES - 1] OF ST_VisuBody;
	p_TempStates						: POINTER TO ARRAY[0..VISU_GlobalConst_Param.VISU_un_MAX_BODIES - 1] OF ST_VisuBodyState;
	p_TempTimestamp						: POINTER TO ULINT;
	p_TempFault							: POINTER TO ST_VisuFault;
END_VAR
m_SetPose := FALSE;
m_Parts(vo_p_Pose => p_TempPose, vo_p_OriginShift => p_TempShift, vo_p_BodyCount => p_TempCount,
	vo_p_Bodies => p_TempBodies, vo_p_BodyStates => p_TempStates, vo_p_Timestamp => p_TempTimestamp,
	vo_p_Fault => p_TempFault);
IF p_TempPose = 0 THEN
	RETURN;
END_IF
(* ST_VisuPose holds LREALs only, so a memory compare sees no padding. *)
m_SetPose := Tc2_System.MEMCMP(ADR(vi_Pose), p_TempPose, SIZEOF(vi_Pose)) <> 0;
IF m_SetPose THEN
	p_TempPose^ := vi_Pose;
	m_NotifyConfigChanged();
END_IF
END_METHOD

END_FUNCTION_BLOCK

// POUs/_FB_VisuVision
(****************************************************************************************************<br>
© Syntegon Group.<br>
All rights reserved, also regarding any disposal, exploitation, reproduction, editing, distribution,<br>
as well as in the event of applications for industrial property rights.<br>
*****************************************************************************************************<br>
DESCRIPTION:<br>
One visualised vision system: a camera over a conveyor. Typical cycle:<br>
  fb_Vision.m_Register(vio_Manifest := GVL_Visu.stManifest, vi_udn_Id := 60, vi_str_Name := 'Vision 1');<br>
  fb_Vision.m_Configure(vi_Pose := LensPose, vi_lr_FieldLength := 400, vi_lr_FieldWidth := 300,<br>
      vi_lr_WorkingDistance := 800);<br>
  fb_Vision.m_SetZone(vi_un_Zone := 1, vi_udn_ConveyorId := 1, vi_lr_Start := 800, vi_lr_End := 1200,<br>
      vi_lr_AllocationOffset := 0, vi_lr_CcsOffset := 1000, vi_lr_StartY := 0, vi_lr_EndY := 0);<br>
  fb_Infeed.m_LatchProduct(..., vi_udn_ClientId := fb_Vision.m_Id());<br>
The pose is the lens, looking along its local -Z. m_Configure describes bodies 1 to 3 (housing, lens,<br>
field of view down to the working distance); further bodies may be added with m_SetBody.<br>
*****************************************************************************************************<br>
VERSION         ¦ DATE       ¦ NAME      ¦ CHANGE<br>
Syn_Visu 4.0.0  ¦ 2026-11-01 ¦ J.Willner ¦ New<br>
****************************************************************************************************)
FUNCTION_BLOCK _FB_VisuVision EXTENDS _FB_VisuDetector

(****************************************************************************************************<br>
© Syntegon Group.<br>
All rights reserved, also regarding any disposal, exploitation, reproduction, editing, distribution,<br>
as well as in the event of applications for industrial property rights.<br>
*****************************************************************************************************<br>
DESCRIPTION:<br>
Manifest type: vision system.<br>
****************************************************************************************************)
METHOD PROTECTED m_ComponentType : E_VisuComponentType
m_ComponentType := E_VisuComponentType.VISION;
END_METHOD

(****************************************************************************************************<br>
© Syntegon Group.<br>
All rights reserved, also regarding any disposal, exploitation, reproduction, editing, distribution,<br>
as well as in the event of applications for industrial property rights.<br>
*****************************************************************************************************<br>
DESCRIPTION:<br>
Sets the lens pose and describes bodies 1 to 3: the housing above the lens, the lens and the field of<br>
view, a frustum from the lens down to the working distance, vi_lr_FieldLength x vi_lr_FieldWidth there.<br>
TRUE if anything changed.<br>
****************************************************************************************************)
METHOD m_Configure : BOOL
VAR_INPUT
	vi_Pose								: ST_VisuPose;	// MCS, the lens looking along its local -Z
	vi_lr_FieldLength					: LREAL;	// [mm] field of view at the working distance, along the local X
	vi_lr_FieldWidth					: LREAL;	// [mm] field of view at the working distance, along the local Y
	vi_lr_WorkingDistance				: LREAL;	// [mm] from the lens to the field of view, e.g. the belt surface
END_VAR
VAR
	TempBefore							: ST_VisuDetectorConfig;
	TempPose							: ST_VisuPose;
	lr_TempDistance						: LREAL;
END_VAR
VAR CONSTANT
	lr_HOUSING_LENGTH					: LREAL := 100;	// [mm]
	lr_HOUSING_WIDTH					: LREAL := 80;	// [mm]
	lr_HOUSING_HEIGHT					: LREAL := 140;	// [mm]
	lr_LENS_DIAMETER					: LREAL := 50;	// [mm]
	lr_LENS_LENGTH						: LREAL := 60;	// [mm]
END_VAR
TempBefore := vo_Visu.stConfig;
lr_TempDistance := MAX(vi_lr_WorkingDistance, 0);
m_SetPose(vi_Pose);
TempPose.fZ := lr_LENS_LENGTH;
m_SetBody(vi_un_Body := 1, vi_e_Shape := E_VisuBodyShape.BOX, vi_e_Role := E_VisuBodyRole.STRUCTURE, vi_Pose := TempPose,
	vi_lr_Length := lr_HOUSING_LENGTH, vi_lr_Width := lr_HOUSING_WIDTH, vi_lr_Height := lr_HOUSING_HEIGHT,
	vi_lr_TopLength := 0, vi_lr_TopWidth := 0);
TempPose.fZ := 0;
m_SetBody(vi_un_Body := 2, vi_e_Shape := E_VisuBodyShape.CYLINDER, vi_e_Role := E_VisuBodyRole.SENSOR, vi_Pose := TempPose,
	vi_lr_Length := lr_LENS_DIAMETER, vi_lr_Width := lr_LENS_DIAMETER, vi_lr_Height := lr_LENS_LENGTH,
	vi_lr_TopLength := 0, vi_lr_TopWidth := 0);
TempPose.fZ := -lr_TempDistance;
m_SetBody(vi_un_Body := 3, vi_e_Shape := E_VisuBodyShape.FRUSTUM, vi_e_Role := E_VisuBodyRole.FIELD_OF_VIEW,
	vi_Pose := TempPose, vi_lr_Length := vi_lr_FieldLength, vi_lr_Width := vi_lr_FieldWidth,
	vi_lr_Height := lr_TempDistance, vi_lr_TopLength := lr_LENS_DIAMETER, vi_lr_TopWidth := lr_LENS_DIAMETER);
m_Configure := Tc2_System.MEMCMP(ADR(TempBefore), ADR(vo_Visu.stConfig), SIZEOF(TempBefore)) <> 0;
END_METHOD

END_FUNCTION_BLOCK

// POUs/_FB_VisuDetector
(****************************************************************************************************<br>
© Syntegon Group.<br>
All rights reserved, also regarding any disposal, exploitation, reproduction, editing, distribution,<br>
as well as in the event of applications for industrial property rights.<br>
*****************************************************************************************************<br>
DESCRIPTION:<br>
Base of a detector (_FB_VisuVision, _FB_VisuSensor): a component that detects products in its zones<br>
and is drawn from the bodies it describes (m_SetBody of _FB_VisuBodyComponent), so the visualisation<br>
needs no code of its own for it. The application latches the products on the conveyor itself<br>
(_FB_VisuConveyor.m_LatchProduct with vi_udn_ClientId := this detector's id). m_Register, called every<br>
cycle, also stamps the state. Not used directly.<br>
*****************************************************************************************************<br>
OUTPUT VALUES:<br>
vo_Visu is the contract structure the gateway reads at the path given to m_Register. Do not write it.<br>
*****************************************************************************************************<br>
VERSION         ¦ DATE       ¦ NAME      ¦ CHANGE<br>
Syn_Visu 4.0.0  ¦ 2026-11-01 ¦ J.Willner ¦ New<br>
Syn_Visu 6.0.0  ¦ 2026-11-01 ¦ J.Willner ¦ Body handling moved to the base _FB_VisuBodyComponent<br>
****************************************************************************************************)
FUNCTION_BLOCK ABSTRACT _FB_VisuDetector EXTENDS _FB_VisuBodyComponent
VAR_OUTPUT
	vo_Visu								: ST_VisuDetector;	// contract structure read by the gateway
END_VAR

(****************************************************************************************************<br>
© Syntegon Group.<br>
All rights reserved, also regarding any disposal, exploitation, reproduction, editing, distribution,<br>
as well as in the event of applications for industrial property rights.<br>
*****************************************************************************************************<br>
DESCRIPTION:<br>
The detector's pose, origin shift, bodies, body states, timestamp and fault for _FB_VisuBodyComponent.<br>
****************************************************************************************************)
METHOD PROTECTED m_Parts : BOOL
VAR_OUTPUT
	vo_p_Pose							: POINTER TO ST_VisuPose;
	vo_p_OriginShift					: POINTER TO ST_VisuPosition;
	vo_p_BodyCount						: POINTER TO UINT;
	vo_p_Bodies							: POINTER TO ARRAY[0..VISU_GlobalConst_Param.VISU_un_MAX_BODIES - 1] OF ST_VisuBody;
	vo_p_BodyStates						: POINTER TO ARRAY[0..VISU_GlobalConst_Param.VISU_un_MAX_BODIES - 1] OF ST_VisuBodyState;
	vo_p_Timestamp						: POINTER TO ULINT;
	vo_p_Fault							: POINTER TO ST_VisuFault;
END_VAR
vo_p_Pose := ADR(vo_Visu.stConfig.stPose);
vo_p_OriginShift := ADR(vo_Visu.stConfig.stOriginShift);
vo_p_BodyCount := ADR(vo_Visu.stConfig.nBodyCount);
vo_p_Bodies := ADR(vo_Visu.stConfig.aBodies);
vo_p_BodyStates := ADR(vo_Visu.stState.aBodyStates);
vo_p_Timestamp := ADR(vo_Visu.stState.nTimestamp);
vo_p_Fault := ADR(vo_Visu.stState.stFault);
m_Parts := TRUE;
END_METHOD

(****************************************************************************************************<br>
© Syntegon Group.<br>
All rights reserved, also regarding any disposal, exploitation, reproduction, editing, distribution,<br>
as well as in the event of applications for industrial property rights.<br>
*****************************************************************************************************<br>
DESCRIPTION:<br>
The detector's zones for _FB_VisuZoneComponent.m_SetZone and m_ClearZones.<br>
****************************************************************************************************)
METHOD PROTECTED m_Zones : BOOL
VAR_OUTPUT
	vo_p_Count							: POINTER TO UINT;
	vo_p_Zones							: POINTER TO ARRAY[0..VISU_GlobalConst_Param.VISU_un_MAX_ZONES - 1] OF ST_VisuZone;
END_VAR
vo_p_Count := ADR(vo_Visu.stConfig.nZoneCount);
vo_p_Zones := ADR(vo_Visu.stConfig.aZones);
m_Zones := TRUE;
END_METHOD

END_FUNCTION_BLOCK

// POUs/_FB_VisuSensor
(****************************************************************************************************<br>
© Syntegon Group.<br>
All rights reserved, also regarding any disposal, exploitation, reproduction, editing, distribution,<br>
as well as in the event of applications for industrial property rights.<br>
*****************************************************************************************************<br>
DESCRIPTION:<br>
One visualised product sensor, e.g. a light barrier at the side of a conveyor. Typical cycle:<br>
  fb_Sensor.m_Register(vio_Manifest := GVL_Visu.stManifest, vi_udn_Id := 61, vi_str_Name := 'Sensor 1');<br>
  fb_Sensor.m_Configure(vi_Pose := HeadPose, vi_lr_BeamLength := 500);<br>
  fb_Sensor.m_SetZone(vi_un_Zone := 1, vi_udn_ConveyorId := 1, vi_lr_Start := 500, vi_lr_End := 500,<br>
      vi_lr_AllocationOffset := 0, vi_lr_CcsOffset := 500, vi_lr_StartY := 0, vi_lr_EndY := 0);<br>
  fb_Sensor.m_SetSignal(vi_b_Signal := b_BeamInterrupted);<br>
The pose is the sensor head; its beam runs along the local +Y. m_Configure describes body 1 (head) and<br>
body 2 (beam); further bodies may be added with m_SetBody.<br>
*****************************************************************************************************<br>
VERSION         ¦ DATE       ¦ NAME      ¦ CHANGE<br>
Syn_Visu 4.0.0  ¦ 2026-11-01 ¦ J.Willner ¦ New<br>
****************************************************************************************************)
FUNCTION_BLOCK _FB_VisuSensor EXTENDS _FB_VisuDetector

(****************************************************************************************************<br>
© Syntegon Group.<br>
All rights reserved, also regarding any disposal, exploitation, reproduction, editing, distribution,<br>
as well as in the event of applications for industrial property rights.<br>
*****************************************************************************************************<br>
DESCRIPTION:<br>
Manifest type: product sensor.<br>
****************************************************************************************************)
METHOD PROTECTED m_ComponentType : E_VisuComponentType
m_ComponentType := E_VisuComponentType.SENSOR;
END_METHOD

(****************************************************************************************************<br>
© Syntegon Group.<br>
All rights reserved, also regarding any disposal, exploitation, reproduction, editing, distribution,<br>
as well as in the event of applications for industrial property rights.<br>
*****************************************************************************************************<br>
DESCRIPTION:<br>
Sets the head pose and describes body 1, the head, and body 2, the beam: a thin cylinder from the head<br>
along its local +Y, vi_lr_BeamLength long. TRUE if anything changed.<br>
****************************************************************************************************)
METHOD m_Configure : BOOL
VAR_INPUT
	vi_Pose								: ST_VisuPose;	// MCS, centre of the head; the beam runs along its local +Y
	vi_lr_BeamLength					: LREAL;	// [mm] e.g. across the belt to the reflector
END_VAR
VAR
	TempBefore							: ST_VisuDetectorConfig;
	TempPose							: ST_VisuPose;
END_VAR
VAR CONSTANT
	lr_HEAD_LENGTH						: LREAL := 30;	// [mm] along the local X
	lr_HEAD_WIDTH						: LREAL := 40;	// [mm] along the local Y, towards the beam
	lr_HEAD_HEIGHT						: LREAL := 60;	// [mm]
	lr_BEAM_DIAMETER					: LREAL := 8;	// [mm]
END_VAR
TempBefore := vo_Visu.stConfig;
m_SetPose(vi_Pose);
TempPose.fZ := -lr_HEAD_HEIGHT / 2;
m_SetBody(vi_un_Body := 1, vi_e_Shape := E_VisuBodyShape.BOX, vi_e_Role := E_VisuBodyRole.SENSOR, vi_Pose := TempPose,
	vi_lr_Length := lr_HEAD_LENGTH, vi_lr_Width := lr_HEAD_WIDTH, vi_lr_Height := lr_HEAD_HEIGHT, vi_lr_TopLength := 0,
	vi_lr_TopWidth := 0);
(* The beam stands on the head's face, turned so that its local +Z runs along the head's +Y. *)
TempPose.fY := lr_HEAD_WIDTH / 2;
TempPose.fZ := 0;
TempPose.fRx := -90;
m_SetBody(vi_un_Body := 2, vi_e_Shape := E_VisuBodyShape.CYLINDER, vi_e_Role := E_VisuBodyRole.BEAM, vi_Pose := TempPose,
	vi_lr_Length := lr_BEAM_DIAMETER, vi_lr_Width := lr_BEAM_DIAMETER, vi_lr_Height := MAX(vi_lr_BeamLength, 0),
	vi_lr_TopLength := 0, vi_lr_TopWidth := 0);
m_Configure := Tc2_System.MEMCMP(ADR(TempBefore), ADR(vo_Visu.stConfig), SIZEOF(TempBefore)) <> 0;
END_METHOD

(****************************************************************************************************<br>
© Syntegon Group.<br>
All rights reserved, also regarding any disposal, exploitation, reproduction, editing, distribution,<br>
as well as in the event of applications for industrial property rights.<br>
*****************************************************************************************************<br>
DESCRIPTION:<br>
Reports the sensor's signal: while TRUE, e.g. while a product interrupts the beam, the beam lights up.<br>
Call once per cycle; it also stamps the state with the cycle's DC time. TRUE.<br>
****************************************************************************************************)
METHOD m_SetSignal : BOOL
VAR_INPUT
	vi_b_Signal							: BOOL;
END_VAR
m_SetSignal := m_SetBodyActive(vi_un_Body := 2, vi_b_Active := vi_b_Signal);
END_METHOD

END_FUNCTION_BLOCK

// POUs/_FB_VisuConveyor
(****************************************************************************************************<br>
© Syntegon Group.<br>
All rights reserved, also regarding any disposal, exploitation, reproduction, editing, distribution,<br>
as well as in the event of applications for industrial property rights.<br>
*****************************************************************************************************<br>
DESCRIPTION:<br>
One visualised conveyor. Typical cycle:<br>
  fb_Infeed.m_Register(vio_Manifest := GVL_Visu.stManifest, vi_udn_Id := 1, vi_str_Name := 'Infeed');<br>
  fb_Infeed.m_Configure(vi_Pose := BeltPose, vi_lr_Length := 5000, vi_lr_Width := 400);<br>
  fb_Infeed.m_SetProductType(vi_udn_Id := 1, vi_lr_Length := 120, vi_lr_Width := 80, vi_lr_Height := 40,<br>
      vi_e_Shape := E_VisuProductShape.BOX, vi_lr_CornerRadius := 0);<br>
  fb_Infeed.m_SetBeltPosition(lr_AxisPosition);  // or m_SetModuloBeltPosition for a modulo axis<br>
  IF b_Latched THEN fb_Infeed.m_LatchProduct(vi_udn_Id := udn_NextId, vi_LatchPose := LatchPose, vi_udn_ProductType := 1,<br>
      vi_lr_LatchBeltPosition := 0, vi_b_UseLatchBeltPosition := FALSE, vi_e_State := E_VisuProductState.DETECTED,<br>
      vi_udn_ClientId := 0); END_IF<br>
m_Configure and m_SetProductType may be called every cycle; the config version only changes when a value does.<br>
*****************************************************************************************************<br>
OUTPUT VALUES:<br>
vo_Visu is the contract structure the gateway reads at the path given to m_Register. Do not write it.<br>
*****************************************************************************************************<br>
VERSION         ¦ DATE       ¦ NAME      ¦ CHANGE<br>
Syn_Visu 3.0.0  ¦ 2026-10-31 ¦ J.Willner ¦ Naming and layout after the TCAT programming guideline<br>
Syn_Visu 3.4.0  ¦ 2026-11-01 ¦ J.Willner ¦ m_LatchProduct: product state and robot (PLACED onto outfeeds)<br>
Syn_Visu 3.5.0  ¦ 2026-11-01 ¦ J.Willner ¦ m_SetProductType: shape and corner radius (protocol 10)<br>
Syn_Visu 4.0.0  ¦ 2026-11-01 ¦ J.Willner ¦ m_LatchProduct: detector that latched the product (protocol 11)<br>
Syn_Visu 7.2.0  ¦ 2026-11-05 ¦ J.Willner ¦ Product index by id; registers rearranged with MEMMOVE<br>
****************************************************************************************************)
FUNCTION_BLOCK _FB_VisuConveyor EXTENDS _FB_VisuComponent
VAR_OUTPUT
	vo_Visu								: ST_VisuConveyor;	// contract structure read by the gateway
END_VAR
VAR
	lr_LastModuloPosition				: LREAL;	// [mm] modulo position of the previous cycle
	b_ModuloInitialised					: BOOL;
	(* Product index: per slot the register index + 1 of a product whose id hashes there, 0 = free. Rebuilt by
	   m_FindProduct after the register was rearranged; m_LatchProduct adds to it. *)
	un_IndexSlot						: ARRAY[0..VISU_GlobalConst_Param.VISU_un_PRODUCT_INDEX_SIZE - 1] OF UINT;
	un_IndexedCount						: UINT;	// [-] register entries the index holds
	b_IndexValid						: BOOL;	// the index matches the register
	b_IndexFailed						: BOOL;	// the index is too small for the register: search linearly
END_VAR

(****************************************************************************************************<br>
© Syntegon Group.<br>
All rights reserved, also regarding any disposal, exploitation, reproduction, editing, distribution,<br>
as well as in the event of applications for industrial property rights.<br>
*****************************************************************************************************<br>
DESCRIPTION:<br>
Takes over vio_New and increments the config version if it differs from the current config. TRUE if changed.<br>
****************************************************************************************************)
METHOD PRIVATE m_ApplyConfig : BOOL
VAR_IN_OUT
	vio_New								: ST_VisuConveyorConfig;
END_VAR
m_ApplyConfig := Tc2_System.MEMCMP(ADR(vio_New), ADR(vo_Visu.stConfig), SIZEOF(vio_New)) <> 0;
IF m_ApplyConfig THEN
	vo_Visu.stConfig := vio_New;
	m_NotifyConfigChanged();
END_IF
END_METHOD

(****************************************************************************************************<br>
© Syntegon Group.<br>
All rights reserved, also regarding any disposal, exploitation, reproduction, editing, distribution,<br>
as well as in the event of applications for industrial property rights.<br>
*****************************************************************************************************<br>
DESCRIPTION:<br>
Belt position last set, [mm].<br>
****************************************************************************************************)
METHOD m_BeltPosition : LREAL
m_BeltPosition := vo_Visu.stState.fBeltPosition;
END_METHOD

(****************************************************************************************************<br>
© Syntegon Group.<br>
All rights reserved, also regarding any disposal, exploitation, reproduction, editing, distribution,<br>
as well as in the event of applications for industrial property rights.<br>
*****************************************************************************************************<br>
DESCRIPTION:<br>
Manifest type: conveyor.<br>
****************************************************************************************************)
METHOD PROTECTED m_ComponentType : E_VisuComponentType
m_ComponentType := E_VisuComponentType.CONVEYOR;
END_METHOD

(****************************************************************************************************<br>
© Syntegon Group.<br>
All rights reserved, also regarding any disposal, exploitation, reproduction, editing, distribution,<br>
as well as in the event of applications for industrial property rights.<br>
*****************************************************************************************************<br>
DESCRIPTION:<br>
Sets pose and size. TRUE if anything changed.<br>
****************************************************************************************************)
METHOD m_Configure : BOOL
VAR_INPUT
	vi_Pose								: ST_VisuPose;	// MCS, belt start on the belt surface; local +X = conveying direction
	vi_lr_Length						: LREAL;	// [mm]
	vi_lr_Width							: LREAL;	// [mm]
END_VAR
VAR
	TempNew								: ST_VisuConveyorConfig;
END_VAR
TempNew := vo_Visu.stConfig;
TempNew.stPose := vi_Pose;
TempNew.fLength := vi_lr_Length;
TempNew.fWidth := vi_lr_Width;
m_Configure := m_ApplyConfig(TempNew);
END_METHOD

(****************************************************************************************************<br>
© Syntegon Group.<br>
All rights reserved, also regarding any disposal, exploitation, reproduction, editing, distribution,<br>
as well as in the event of applications for industrial property rights.<br>
*****************************************************************************************************<br>
DESCRIPTION:<br>
Register index of the product with vi_udn_Id, -1 if not found. Looks it up in the product index by id, which it<br>
rebuilds first after the register was rearranged; searches linearly only if the index is too small.<br>
****************************************************************************************************)
METHOD m_FindProduct : INT
VAR_INPUT
	vi_udn_Id							: UDINT;	// [-] product id
END_VAR
VAR
	un_TempIndex						: UINT;
	un_TempSlot							: UINT;
	un_TempProbe						: UINT;
	un_TempEntry						: UINT;	// [-] register index + 1, 0 = free slot
END_VAR
m_FindProduct := -1;
IF NOT b_IndexFailed AND (NOT b_IndexValid OR un_IndexedCount <> vo_Visu.stState.nProductCount) THEN
	m_IndexRebuild();
END_IF

IF b_IndexValid THEN
	un_TempSlot := m_IndexSlotOf(vi_udn_Id);
	FOR un_TempProbe := 1 TO VISU_GlobalConst_Param.VISU_un_PRODUCT_INDEX_SIZE DO
		un_TempEntry := un_IndexSlot[un_TempSlot];
		IF un_TempEntry = 0 THEN
			RETURN;
		END_IF
		IF un_TempEntry <= vo_Visu.stState.nProductCount THEN
			IF vo_Visu.stState.aProducts[un_TempEntry - 1].nId = vi_udn_Id THEN
				m_FindProduct := UINT_TO_INT(un_TempEntry - 1);
				RETURN;
			END_IF
		END_IF
		un_TempSlot := (un_TempSlot + 1) AND (VISU_GlobalConst_Param.VISU_un_PRODUCT_INDEX_SIZE - 1);
	END_FOR
	RETURN;
END_IF

(* Index too small for the register: search linearly. *)
un_TempIndex := 0;
WHILE un_TempIndex < vo_Visu.stState.nProductCount DO
	IF vo_Visu.stState.aProducts[un_TempIndex].nId = vi_udn_Id THEN
		m_FindProduct := UINT_TO_INT(un_TempIndex);
		RETURN;
	END_IF
	un_TempIndex := un_TempIndex + 1;
END_WHILE
END_METHOD

(****************************************************************************************************<br>
© Syntegon Group.<br>
All rights reserved, also regarding any disposal, exploitation, reproduction, editing, distribution,<br>
as well as in the event of applications for industrial property rights.<br>
*****************************************************************************************************<br>
DESCRIPTION:<br>
Reads register entry vi_un_Index and its current pose in the conveyor's coordinate system (latch pose moved<br>
along the belt by the belt travel since).<br>
Indices shift when products are removed; use the product id to follow a product.<br>
*****************************************************************************************************<br>
OUTPUT VALUES:<br>
FALSE if vi_un_Index is out of range.<br>
****************************************************************************************************)
METHOD m_GetProduct : BOOL
VAR_INPUT
	vi_un_Index							: UINT;	// [-] 0..m_ProductCount() - 1
END_VAR
VAR_OUTPUT
	vo_Product							: ST_VisuProduct;
	vo_Pose								: ST_VisuPlanarPose;	// conveyor coordinate system, current bottom centre
END_VAR
m_GetProduct := vi_un_Index < vo_Visu.stState.nProductCount;
IF m_GetProduct THEN
	vo_Product := vo_Visu.stState.aProducts[vi_un_Index];
	vo_Pose := m_ProductPose(vo_Product);
END_IF
END_METHOD

(****************************************************************************************************<br>
© Syntegon Group.<br>
All rights reserved, also regarding any disposal, exploitation, reproduction, editing, distribution,<br>
as well as in the event of applications for industrial property rights.<br>
*****************************************************************************************************<br>
DESCRIPTION:<br>
Adds register entry vi_un_Index with product id vi_udn_Id to the product index, in the first free slot from<br>
its hash slot on.<br>
*****************************************************************************************************<br>
OUTPUT VALUES:<br>
FALSE if the index has no free slot (VISU_un_PRODUCT_INDEX_SIZE too small for VISU_un_MAX_PRODUCTS).<br>
****************************************************************************************************)
METHOD PRIVATE m_IndexInsert : BOOL
VAR_INPUT
	vi_udn_Id							: UDINT;	// [-] product id
	vi_un_Index							: UINT;	// [-] register index
END_VAR
VAR
	un_TempSlot							: UINT;
	un_TempProbe						: UINT;
END_VAR
m_IndexInsert := FALSE;
un_TempSlot := m_IndexSlotOf(vi_udn_Id);
FOR un_TempProbe := 1 TO VISU_GlobalConst_Param.VISU_un_PRODUCT_INDEX_SIZE DO
	IF un_IndexSlot[un_TempSlot] = 0 THEN
		un_IndexSlot[un_TempSlot] := vi_un_Index + 1;
		m_IndexInsert := TRUE;
		RETURN;
	END_IF
	un_TempSlot := (un_TempSlot + 1) AND (VISU_GlobalConst_Param.VISU_un_PRODUCT_INDEX_SIZE - 1);
END_FOR
END_METHOD

(****************************************************************************************************<br>
© Syntegon Group.<br>
All rights reserved, also regarding any disposal, exploitation, reproduction, editing, distribution,<br>
as well as in the event of applications for industrial property rights.<br>
*****************************************************************************************************<br>
DESCRIPTION:<br>
Builds the product index from the register anew, e.g. after products were removed and the register moved up.<br>
If the index is too small for the register, it gives up for good and m_FindProduct searches linearly.<br>
*****************************************************************************************************<br>
OUTPUT VALUES:<br>
TRUE if the index matches the register.<br>
****************************************************************************************************)
METHOD PRIVATE m_IndexRebuild : BOOL
VAR
	un_TempIndex						: UINT;
END_VAR
Tc2_System.MEMSET(ADR(un_IndexSlot), 0, SIZEOF(un_IndexSlot));
b_IndexValid := TRUE;
un_TempIndex := 0;
WHILE un_TempIndex < vo_Visu.stState.nProductCount DO
	IF NOT m_IndexInsert(vo_Visu.stState.aProducts[un_TempIndex].nId, un_TempIndex) THEN
		b_IndexValid := FALSE;
		b_IndexFailed := TRUE;
		EXIT;
	END_IF
	un_TempIndex := un_TempIndex + 1;
END_WHILE
un_IndexedCount := vo_Visu.stState.nProductCount;
m_IndexRebuild := b_IndexValid;
END_METHOD

(****************************************************************************************************<br>
© Syntegon Group.<br>
All rights reserved, also regarding any disposal, exploitation, reproduction, editing, distribution,<br>
as well as in the event of applications for industrial property rights.<br>
*****************************************************************************************************<br>
DESCRIPTION:<br>
First slot of the product index to look at for a product id (multiplicative hash): consecutive ids land on<br>
different slots. The search goes on slot by slot from there.<br>
****************************************************************************************************)
METHOD PRIVATE m_IndexSlotOf : UINT
VAR_INPUT
	vi_udn_Id							: UDINT;	// [-] product id
END_VAR
(* The product wraps around in 32 bits on purpose. *)
m_IndexSlotOf := UDINT_TO_UINT((vi_udn_Id * UDINT#2654435761) AND UINT_TO_UDINT(VISU_GlobalConst_Param.VISU_un_PRODUCT_INDEX_SIZE - 1));
END_METHOD

(****************************************************************************************************<br>
© Syntegon Group.<br>
All rights reserved, also regarding any disposal, exploitation, reproduction, editing, distribution,<br>
as well as in the event of applications for industrial property rights.<br>
*****************************************************************************************************<br>
DESCRIPTION:<br>
Adds a product at the current belt position. Call m_SetBeltPosition first in the cycle,<br>
or pass the belt position at the latch moment in vi_lr_LatchBeltPosition.<br>
A product arriving on the conveyor enters as DETECTED (default), naming the client that latched it (vision<br>
system, sensor, station). A product a robot puts down onto it (outfeed, tray, back onto the same belt)<br>
enters as PLACED with that robot as client: the visualisation shows a DETECTED or ASSIGNED product passing<br>
the belt end as missed. Its previous state is the state it enters in.<br>
*****************************************************************************************************<br>
OUTPUT VALUES:<br>
FALSE for vi_udn_Id = 0, an id already in the register, or a full register.<br>
****************************************************************************************************)
METHOD m_LatchProduct : BOOL
VAR_INPUT
	vi_udn_Id							: UDINT;	// [-] unique on this conveyor, > 0
	vi_LatchPose						: ST_VisuPlanarPose;	// conveyor coordinate system (from its origin shift), bottom centre at the latch moment
	vi_udn_ProductType					: UDINT;	// [-] id given to m_SetProductType
	vi_lr_LatchBeltPosition				: LREAL;	// [mm] used only if vi_b_UseLatchBeltPosition, else 0
	vi_b_UseLatchBeltPosition			: BOOL;	// FALSE: latch at the current belt position
	vi_e_State							: E_VisuProductState;	// DETECTED for a product arriving, PLACED for a product put down by a robot
	vi_udn_ClientId						: UDINT;	// [-] manifest id of the client that latched it or put it down, 0 = none
END_VAR
VAR
	un_TempIndex						: UINT;
END_VAR
m_LatchProduct := FALSE;
un_TempIndex := vo_Visu.stState.nProductCount;
IF vi_udn_Id = 0 OR m_FindProduct(vi_udn_Id) >= 0 OR un_TempIndex >= VISU_GlobalConst_Param.VISU_un_MAX_PRODUCTS THEN
	RETURN;
END_IF
vo_Visu.stState.aProducts[un_TempIndex].nId := vi_udn_Id;
vo_Visu.stState.aProducts[un_TempIndex].bValid := TRUE;
vo_Visu.stState.aProducts[un_TempIndex].stLatchPose := vi_LatchPose;
IF vi_b_UseLatchBeltPosition THEN
	vo_Visu.stState.aProducts[un_TempIndex].fLatchBeltPosition := vi_lr_LatchBeltPosition;
ELSE
	vo_Visu.stState.aProducts[un_TempIndex].fLatchBeltPosition := vo_Visu.stState.fBeltPosition;
END_IF
vo_Visu.stState.aProducts[un_TempIndex].eState := vi_e_State;
vo_Visu.stState.aProducts[un_TempIndex].ePreviousState := vi_e_State;
vo_Visu.stState.aProducts[un_TempIndex].nLastClientId := vi_udn_ClientId;
vo_Visu.stState.aProducts[un_TempIndex].nMoverId := 0;
vo_Visu.stState.aProducts[un_TempIndex].nFingerId := 0;
vo_Visu.stState.aProducts[un_TempIndex].nProductType := vi_udn_ProductType;
vo_Visu.stState.nProductCount := un_TempIndex + 1;
(* m_FindProduct above brought the index up to the register; the new entry joins it. *)
IF b_IndexValid AND un_IndexedCount = un_TempIndex THEN
	IF m_IndexInsert(vi_udn_Id, un_TempIndex) THEN
		un_IndexedCount := un_TempIndex + 1;
	ELSE
		b_IndexValid := FALSE;
		b_IndexFailed := TRUE;
	END_IF
END_IF
vo_Visu.stState.nTimestamp := m_DcTime();
m_LatchProduct := TRUE;
END_METHOD

(****************************************************************************************************<br>
© Syntegon Group.<br>
All rights reserved, also regarding any disposal, exploitation, reproduction, editing, distribution,<br>
as well as in the event of applications for industrial property rights.<br>
*****************************************************************************************************<br>
DESCRIPTION:<br>
Puts a product of the register at a new pose (conveyor coordinate system) at the current belt position, e.g. while a mover pushes it<br>
along the belt faster than the belt runs. Call m_SetBeltPosition first in the cycle. Keeps its state.<br>
*****************************************************************************************************<br>
OUTPUT VALUES:<br>
FALSE if the product is not in the register.<br>
****************************************************************************************************)
METHOD m_MoveProduct : BOOL
VAR_INPUT
	vi_udn_Id							: UDINT;	// [-] product id
	vi_Pose								: ST_VisuPlanarPose;	// conveyor coordinate system, bottom centre of the product now
END_VAR
VAR
	n_TempIndex							: INT;
END_VAR
n_TempIndex := m_FindProduct(vi_udn_Id);
m_MoveProduct := n_TempIndex >= 0;
IF m_MoveProduct THEN
	vo_Visu.stState.aProducts[n_TempIndex].stLatchPose := vi_Pose;
	vo_Visu.stState.aProducts[n_TempIndex].fLatchBeltPosition := vo_Visu.stState.fBeltPosition;
	vo_Visu.stState.nTimestamp := m_DcTime();
END_IF
END_METHOD

(****************************************************************************************************<br>
© Syntegon Group.<br>
All rights reserved, also regarding any disposal, exploitation, reproduction, editing, distribution,<br>
as well as in the event of applications for industrial property rights.<br>
*****************************************************************************************************<br>
DESCRIPTION:<br>
Number of products in the register; valid indices for m_GetProduct are 0..m_ProductCount() - 1.<br>
****************************************************************************************************)
METHOD m_ProductCount : UINT
m_ProductCount := vo_Visu.stState.nProductCount;
END_METHOD

(****************************************************************************************************<br>
© Syntegon Group.<br>
All rights reserved, also regarding any disposal, exploitation, reproduction, editing, distribution,<br>
as well as in the event of applications for industrial property rights.<br>
*****************************************************************************************************<br>
DESCRIPTION:<br>
Current pose of a product in the conveyor's coordinate system: latch pose moved along the belt<br>
(local +X) by the belt travel since the latch.<br>
****************************************************************************************************)
METHOD PRIVATE m_ProductPose : ST_VisuPlanarPose
VAR_IN_OUT CONSTANT
	vio_Product							: ST_VisuProduct;
END_VAR
VAR
	lr_TempTravel						: LREAL;	// [mm]
END_VAR
lr_TempTravel := vo_Visu.stState.fBeltPosition - vio_Product.fLatchBeltPosition;
m_ProductPose := vio_Product.stLatchPose;
m_ProductPose.fX := m_ProductPose.fX + lr_TempTravel;
END_METHOD

(****************************************************************************************************<br>
© Syntegon Group.<br>
All rights reserved, also regarding any disposal, exploitation, reproduction, editing, distribution,<br>
as well as in the event of applications for industrial property rights.<br>
*****************************************************************************************************<br>
DESCRIPTION:<br>
Removes a product from the register. FALSE if it is not in the register.<br>
****************************************************************************************************)
METHOD m_RemoveProduct : BOOL
VAR_INPUT
	vi_udn_Id							: UDINT;	// [-] product id
END_VAR
VAR
	n_TempIndex							: INT;
	n_TempLast							: INT;
END_VAR
n_TempIndex := m_FindProduct(vi_udn_Id);
m_RemoveProduct := n_TempIndex >= 0;
IF NOT m_RemoveProduct THEN
	RETURN;
END_IF
n_TempLast := UINT_TO_INT(vo_Visu.stState.nProductCount) - 1;
(* The entries behind it move up by one, in one go. *)
IF n_TempIndex < n_TempLast THEN
	Tc2_System.MEMMOVE(ADR(vo_Visu.stState.aProducts[n_TempIndex]), ADR(vo_Visu.stState.aProducts[n_TempIndex + 1]),
		INT_TO_UDINT(n_TempLast - n_TempIndex) * SIZEOF(ST_VisuProduct));
END_IF
vo_Visu.stState.aProducts[n_TempLast].bValid := FALSE;
vo_Visu.stState.nProductCount := INT_TO_UINT(n_TempLast);
b_IndexValid := FALSE;
vo_Visu.stState.nTimestamp := m_DcTime();
END_METHOD

(****************************************************************************************************<br>
© Syntegon Group.<br>
All rights reserved, also regarding any disposal, exploitation, reproduction, editing, distribution,<br>
as well as in the event of applications for industrial property rights.<br>
*****************************************************************************************************<br>
DESCRIPTION:<br>
Housekeeping: drops invalid entries and products that have travelled beyond vi_lr_BeltX (along the<br>
conveyor from its start). Products a robot is working on (ASSIGNED or PICKED) are kept wherever they are.<br>
The entries that stay move up in runs (usually one: the products leaving are the oldest, at the front).<br>
*****************************************************************************************************<br>
OUTPUT VALUES:<br>
Number of removed entries.<br>
****************************************************************************************************)
METHOD m_RemoveProductsBeyond : UINT
VAR_INPUT
	vi_lr_BeltX							: LREAL;	// [mm] e.g. belt length + some margin so missed products stay visible briefly
END_VAR
VAR
	un_TempCount						: UINT;	// [-] entries before
	un_TempRead							: UINT;
	un_TempWrite						: UINT;
	un_TempRunStart						: UINT;	// [-] first entry of a run of entries that stay
	b_TempStays							: BOOL;
END_VAR
m_RemoveProductsBeyond := 0;
un_TempCount := vo_Visu.stState.nProductCount;
IF un_TempCount = 0 THEN
	RETURN;
END_IF

(* Keep the entries that stay, in order, moving each run of them up in one go. *)
un_TempWrite := 0;
un_TempRead := 0;
WHILE un_TempRead < un_TempCount DO
	IF m_StaysInRegister(un_TempRead, vi_lr_BeltX) THEN
		un_TempRunStart := un_TempRead;
		b_TempStays := TRUE;
		WHILE b_TempStays DO
			un_TempRead := un_TempRead + 1;
			b_TempStays := FALSE;
			IF un_TempRead < un_TempCount THEN
				b_TempStays := m_StaysInRegister(un_TempRead, vi_lr_BeltX);
			END_IF
		END_WHILE
		IF un_TempWrite <> un_TempRunStart THEN
			Tc2_System.MEMMOVE(ADR(vo_Visu.stState.aProducts[un_TempWrite]), ADR(vo_Visu.stState.aProducts[un_TempRunStart]),
				UINT_TO_UDINT(un_TempRead - un_TempRunStart) * SIZEOF(ST_VisuProduct));
		END_IF
		un_TempWrite := un_TempWrite + (un_TempRead - un_TempRunStart);
	ELSE
		un_TempRead := un_TempRead + 1;
	END_IF
END_WHILE

(* Invalidate the freed tail. *)
m_RemoveProductsBeyond := un_TempCount - un_TempWrite;
IF un_TempWrite < un_TempCount THEN
	FOR un_TempRead := un_TempWrite TO un_TempCount - 1 DO
		vo_Visu.stState.aProducts[un_TempRead].bValid := FALSE;
	END_FOR
	vo_Visu.stState.nProductCount := un_TempWrite;
	vo_Visu.stState.nTimestamp := m_DcTime();
	b_IndexValid := FALSE;
END_IF
END_METHOD

(****************************************************************************************************<br>
© Syntegon Group.<br>
All rights reserved, also regarding any disposal, exploitation, reproduction, editing, distribution,<br>
as well as in the event of applications for industrial property rights.<br>
*****************************************************************************************************<br>
DESCRIPTION:<br>
Sets the belt position: how far the belt surface has travelled, continuous (no modulo).<br>
Call once per cycle; it also stamps the state with the cycle's DC time.<br>
****************************************************************************************************)
METHOD m_SetBeltPosition : BOOL
VAR_INPUT
	vi_lr_Position						: LREAL;	// [mm]
END_VAR
vo_Visu.stState.fBeltPosition := vi_lr_Position;
vo_Visu.stState.nTimestamp := m_DcTime();
m_SetBeltPosition := TRUE;
END_METHOD

(****************************************************************************************************<br>
© Syntegon Group.<br>
All rights reserved, also regarding any disposal, exploitation, reproduction, editing, distribution,<br>
as well as in the event of applications for industrial property rights.<br>
*****************************************************************************************************<br>
DESCRIPTION:<br>
Sets whether the belt is drawn as a body. A conveyor without one (FALSE) shows only its products, zones and<br>
its axis from the origin to the conveying direction arrow. Default TRUE. TRUE if anything changed.<br>
****************************************************************************************************)
METHOD m_SetBodyVisible : BOOL
VAR_INPUT
	vi_b_Visible						: BOOL;	// TRUE = drawn as a body, FALSE = a conveyor without one
END_VAR
VAR
	TempNew								: ST_VisuConveyorConfig;
END_VAR
TempNew := vo_Visu.stConfig;
TempNew.bBody := vi_b_Visible;
m_SetBodyVisible := m_ApplyConfig(TempNew);
END_METHOD

(****************************************************************************************************<br>
© Syntegon Group.<br>
All rights reserved, also regarding any disposal, exploitation, reproduction, editing, distribution,<br>
as well as in the event of applications for industrial property rights.<br>
*****************************************************************************************************<br>
DESCRIPTION:<br>
Sets or clears the fault of the conveyor: drawn red with the message while active. The fault stays until it<br>
is cleared with m_SetFault(vi_b_Active := FALSE, vi_str_Message := ''). TRUE.<br>
****************************************************************************************************)
METHOD m_SetFault : BOOL
VAR_INPUT
	vi_b_Active							: BOOL;	// TRUE: fault active
	vi_str_Message						: STRING(80);	// shown to the operator; empty shows 'Fault'
END_VAR
vo_Visu.stState.stFault.bActive := vi_b_Active;
vo_Visu.stState.stFault.sMessage := vi_str_Message;
m_SetFault := TRUE;
END_METHOD

(****************************************************************************************************<br>
© Syntegon Group.<br>
All rights reserved, also regarding any disposal, exploitation, reproduction, editing, distribution,<br>
as well as in the event of applications for industrial property rights.<br>
*****************************************************************************************************<br>
DESCRIPTION:<br>
Like m_SetBeltPosition, for a modulo axis: unwraps the position so the belt position stays continuous.<br>
Call once per cycle.<br>
*****************************************************************************************************<br>
LIMITS:<br>
The axis must move less than half a modulo period per cycle.<br>
****************************************************************************************************)
METHOD m_SetModuloBeltPosition : BOOL
VAR_INPUT
	vi_lr_ModuloPosition				: LREAL;	// [mm] in [0, vi_lr_ModuloPeriod)
	vi_lr_ModuloPeriod					: LREAL;	// [mm] <= 0 passes vi_lr_ModuloPosition through unchanged
	vi_b_Reset							: BOOL;	// TRUE: restart the belt position at vi_lr_ModuloPosition
END_VAR
VAR
	lr_TempPosition						: LREAL;	// [mm]
	lr_TempDelta						: LREAL;	// [mm]
END_VAR
IF vi_b_Reset OR NOT b_ModuloInitialised OR vi_lr_ModuloPeriod <= 0 THEN
	lr_TempPosition := vi_lr_ModuloPosition;
	b_ModuloInitialised := TRUE;
ELSE
	lr_TempDelta := vi_lr_ModuloPosition - lr_LastModuloPosition;
	IF lr_TempDelta > vi_lr_ModuloPeriod / 2 THEN
		lr_TempDelta := lr_TempDelta - vi_lr_ModuloPeriod;
	ELSIF lr_TempDelta < -vi_lr_ModuloPeriod / 2 THEN
		lr_TempDelta := lr_TempDelta + vi_lr_ModuloPeriod;
	END_IF
	lr_TempPosition := vo_Visu.stState.fBeltPosition + lr_TempDelta;
END_IF
lr_LastModuloPosition := vi_lr_ModuloPosition;
m_SetModuloBeltPosition := m_SetBeltPosition(lr_TempPosition);
END_METHOD

(****************************************************************************************************<br>
© Syntegon Group.<br>
All rights reserved, also regarding any disposal, exploitation, reproduction, editing, distribution,<br>
as well as in the event of applications for industrial property rights.<br>
*****************************************************************************************************<br>
DESCRIPTION:<br>
Moves the conveyor's coordinate system away from the belt start (stPose), in the belt's local frame. Belt<br>
coordinates (zones' start, end and CCS offset) then count from the shifted origin. TRUE if anything changed.<br>
****************************************************************************************************)
METHOD m_SetOriginShift : BOOL
VAR_INPUT
	vi_lr_X								: LREAL;	// [mm] along the conveying direction
	vi_lr_Y								: LREAL;	// [mm] across the belt, 0 = none
	vi_lr_Z								: LREAL;	// [mm] along the belt surface normal, 0 = none
END_VAR
VAR
	TempNew								: ST_VisuConveyorConfig;
END_VAR
TempNew := vo_Visu.stConfig;
TempNew.stOriginShift.fX := vi_lr_X;
TempNew.stOriginShift.fY := vi_lr_Y;
TempNew.stOriginShift.fZ := vi_lr_Z;
m_SetOriginShift := m_ApplyConfig(TempNew);
END_METHOD

(****************************************************************************************************<br>
© Syntegon Group.<br>
All rights reserved, also regarding any disposal, exploitation, reproduction, editing, distribution,<br>
as well as in the event of applications for industrial property rights.<br>
*****************************************************************************************************<br>
DESCRIPTION:<br>
Changes a product's state and names the client that changed it: the robot that is assigned to, picks,<br>
places or releases it, the station that rejects it. The state before is kept as ePreviousState when the<br>
state changes; calling it again with the same state keeps it. FALSE if the product is not in the register.<br>
****************************************************************************************************)
METHOD m_SetProductState : BOOL
VAR_INPUT
	vi_udn_Id							: UDINT;	// [-] product id
	vi_e_State							: E_VisuProductState;
	vi_udn_ClientId						: UDINT;	// [-] manifest id of the client making the change, 0 = none
	vi_udn_MoverId						: UDINT;	// [-] mover of an XTS gantry or loop carrying the product, 0 = none
	vi_udn_FingerId						: UDINT;	// [-] gripper finger (1-based) the product hangs from while picked, 0 = the flange
END_VAR
VAR
	n_TempIndex							: INT;
END_VAR
n_TempIndex := m_FindProduct(vi_udn_Id);
m_SetProductState := n_TempIndex >= 0;
IF m_SetProductState THEN
	IF vo_Visu.stState.aProducts[n_TempIndex].eState <> vi_e_State THEN
		vo_Visu.stState.aProducts[n_TempIndex].ePreviousState := vo_Visu.stState.aProducts[n_TempIndex].eState;
	END_IF
	vo_Visu.stState.aProducts[n_TempIndex].eState := vi_e_State;
	vo_Visu.stState.aProducts[n_TempIndex].nLastClientId := vi_udn_ClientId;
	vo_Visu.stState.aProducts[n_TempIndex].nMoverId := vi_udn_MoverId;
	vo_Visu.stState.aProducts[n_TempIndex].nFingerId := vi_udn_FingerId;
	vo_Visu.stState.nTimestamp := m_DcTime();
END_IF
END_METHOD

